screen "D_GraphicView_1" 800x480
   GraphicView "Static" at 6,4 size 100x60
   TextField "Label_Static" at 6,96 size 148x16; Text 'Static'
   GraphicView "A_Range" at 158,4 size 100x60
      Appearance <- "D_Range"
   TextField "Label_A_Range" at 158,96 size 148x16; Text 'A_Range'
   GraphicView "A_Flash" at 310,4 size 100x60
      Appearance <- "D_Range"
   TextField "Label_A_Flash" at 310,96 size 148x16; Text 'A_Flash'
   GraphicView "A_Bit" at 462,4 size 100x60
      Appearance <- "D_Bool"
   TextField "Label_A_Bit" at 462,96 size 148x16; Text 'A_Bit'
   GraphicView "A_Bits" at 614,4 size 100x60
      Appearance <- "D_Bits"
   TextField "Label_A_Bits" at 614,96 size 148x16; Text 'A_Bits'
   GraphicView "V_Range" at 6,116 size 100x60
      Visibility <- "D_Range"
   TextField "Label_V_Range" at 6,208 size 148x16; Text 'V_Range'
   GraphicView "V_Bit" at 158,116 size 100x60
      Visibility <- "D_Vis"
   TextField "Label_V_Bit" at 158,208 size 148x16; Text 'V_Bit'
   GraphicView "M_H" at 310,116 size 100x60
      HorizontalMovement <- "D_Pct"
   TextField "Label_M_H" at 310,208 size 148x16; Text 'M_H'
   GraphicView "M_V" at 462,116 size 100x60
      VerticalMovement <- "D_Pct"
   TextField "Label_M_V" at 462,208 size 148x16; Text 'M_V'
   GraphicView "M_D" at 614,116 size 100x60
      DiagonalMovement <- "D_Pct"
   TextField "Label_M_D" at 614,208 size 148x16; Text 'M_D'
   GraphicView "M_Direct" at 6,228 size 100x60
      DirectMovement <- "D_X"
      DirectMovement <- "D_Y"
   TextField "Label_M_Direct" at 6,320 size 148x16; Text 'M_Direct'
   GraphicView "E_Range" at 158,228 size 100x60
      ObjectEnable <- "D_Range"
   TextField "Label_E_Range" at 158,320 size 148x16; Text 'E_Range'
   GraphicView "E_Bit" at 310,228 size 100x60
      ObjectEnable <- "D_En"
   TextField "Label_E_Bit" at 310,320 size 148x16; Text 'E_Bit'
   IOField "State" at 4,454 size 60x22; FormatPattern 9
      ProcessValue <- "D_State"
   Button "S1" at 70,454 size 40x22; TextOff 'S1'
      on Click: "SetS1"()
   Button "S2" at 114,454 size 40x22; TextOff 'S2'
      on Click: "SetS2"()
   Button "S3" at 158,454 size 40x22; TextOff 'S3'
      on Click: "SetS3"()
   Button "S4" at 202,454 size 40x22; TextOff 'S4'
      on Click: "SetS4"()
   Button "Next" at 756,454 size 40x22; TextOff 'Next'
      on Click: ActivateScreen("D_IOField_1", 0)

screen "D_IOField_2" 800x480
   IOField "PV_Int_Output" at 6,4 size 100x30; FormatPattern s99999
      ProcessValue <- "D_Int"
   TextField "Label_PV_Int_Output" at 6,66 size 148x16; Text 'PV_Int_Output'
   IOField "PV_Int_s99" at 158,4 size 100x30; FormatPattern s99
      ProcessValue <- "D_Int"
   TextField "Label_PV_Int_s99" at 158,66 size 148x16; Text 'PV_Int_s99'
   IOField "State" at 4,454 size 60x22; FormatPattern 9
      ProcessValue <- "D_State"
   Button "S1" at 70,454 size 40x22; TextOff 'S1'
      on Click: "SetS1"()
   Button "S2" at 114,454 size 40x22; TextOff 'S2'
      on Click: "SetS2"()
   Button "S3" at 158,454 size 40x22; TextOff 'S3'
      on Click: "SetS3"()
   Button "S4" at 202,454 size 40x22; TextOff 'S4'
      on Click: "SetS4"()
   Button "Next" at 756,454 size 40x22; TextOff 'Next'
      on Click: ActivateScreen("D_Button_1", 0)

screen "D_Line_1" 800x480
   TextField "Label_Static" at 6,86 size 148x16; Text 'Static'
   Line "A_Range" at 158,4 size 100x50
      Appearance <- "D_Range"
   TextField "Label_A_Range" at 158,86 size 148x16; Text 'A_Range'
   Line "A_Flash" at 310,4 size 100x50
      Appearance <- "D_Range"
   TextField "Label_A_Flash" at 310,86 size 148x16; Text 'A_Flash'
   Line "A_Bit" at 462,4 size 100x50
      Appearance <- "D_Bool"
   TextField "Label_A_Bit" at 462,86 size 148x16; Text 'A_Bit'
   Line "A_Bits" at 614,4 size 100x50
      Appearance <- "D_Bits"
   TextField "Label_A_Bits" at 614,86 size 148x16; Text 'A_Bits'
   Line "V_Range" at 6,106 size 100x50
      Visibility <- "D_Range"
   TextField "Label_V_Range" at 6,188 size 148x16; Text 'V_Range'
   Line "V_Bit" at 158,106 size 100x50
      Visibility <- "D_Vis"
   TextField "Label_V_Bit" at 158,188 size 148x16; Text 'V_Bit'
   Line "M_H" at 310,106 size 100x50
      HorizontalMovement <- "D_Pct"
   TextField "Label_M_H" at 310,188 size 148x16; Text 'M_H'
   Line "M_V" at 462,106 size 100x50
      VerticalMovement <- "D_Pct"
   TextField "Label_M_V" at 462,188 size 148x16; Text 'M_V'
   Line "M_D" at 614,106 size 100x50
      DiagonalMovement <- "D_Pct"
   TextField "Label_M_D" at 614,188 size 148x16; Text 'M_D'
   Line "M_Direct" at 6,208 size 100x50
      DirectMovement <- "D_X"
      DirectMovement <- "D_Y"
   TextField "Label_M_Direct" at 6,290 size 148x16; Text 'M_Direct'
   Line "E_Range" at 158,208 size 100x50
      ObjectEnable <- "D_Range"
   TextField "Label_E_Range" at 158,290 size 148x16; Text 'E_Range'
   Line "E_Bit" at 310,208 size 100x50
      ObjectEnable <- "D_En"
   TextField "Label_E_Bit" at 310,290 size 148x16; Text 'E_Bit'
   IOField "State" at 4,454 size 60x22; FormatPattern 9
      ProcessValue <- "D_State"
   Button "S1" at 70,454 size 40x22; TextOff 'S1'
      on Click: "SetS1"()
   Button "S2" at 114,454 size 40x22; TextOff 'S2'
      on Click: "SetS2"()
   Button "S3" at 158,454 size 40x22; TextOff 'S3'
      on Click: "SetS3"()
   Button "S4" at 202,454 size 40x22; TextOff 'S4'
      on Click: "SetS4"()
   Button "Next" at 756,454 size 40x22; TextOff 'Next'
      on Click: ActivateScreen("D_Polyline_1", 0)

screen "D_Polygon_1" 800x480
   TextField "Label_Static" at 6,86 size 148x16; Text 'Static'
   Polygon "A_Range" at 158,4 size 100x50
      Appearance <- "D_Range"
   TextField "Label_A_Range" at 158,86 size 148x16; Text 'A_Range'
   Polygon "A_Flash" at 310,4 size 100x50
      Appearance <- "D_Range"
   TextField "Label_A_Flash" at 310,86 size 148x16; Text 'A_Flash'
   Polygon "A_Bit" at 462,4 size 100x50
      Appearance <- "D_Bool"
   TextField "Label_A_Bit" at 462,86 size 148x16; Text 'A_Bit'
   Polygon "A_Bits" at 614,4 size 100x50
      Appearance <- "D_Bits"
   TextField "Label_A_Bits" at 614,86 size 148x16; Text 'A_Bits'
   Polygon "V_Range" at 6,106 size 100x50
      Visibility <- "D_Range"
   TextField "Label_V_Range" at 6,188 size 148x16; Text 'V_Range'
   Polygon "V_Bit" at 158,106 size 100x50
      Visibility <- "D_Vis"
   TextField "Label_V_Bit" at 158,188 size 148x16; Text 'V_Bit'
   Polygon "M_H" at 310,106 size 100x50
      HorizontalMovement <- "D_Pct"
   TextField "Label_M_H" at 310,188 size 148x16; Text 'M_H'
   Polygon "M_V" at 462,106 size 100x50
      VerticalMovement <- "D_Pct"
   TextField "Label_M_V" at 462,188 size 148x16; Text 'M_V'
   Polygon "M_D" at 614,106 size 100x50
      DiagonalMovement <- "D_Pct"
   TextField "Label_M_D" at 614,188 size 148x16; Text 'M_D'
   Polygon "M_Direct" at 6,208 size 100x50
      DirectMovement <- "D_X"
      DirectMovement <- "D_Y"
   TextField "Label_M_Direct" at 6,290 size 148x16; Text 'M_Direct'
   Polygon "E_Range" at 158,208 size 100x50
      ObjectEnable <- "D_Range"
   TextField "Label_E_Range" at 158,290 size 148x16; Text 'E_Range'
   Polygon "E_Bit" at 310,208 size 100x50
      ObjectEnable <- "D_En"
   TextField "Label_E_Bit" at 310,290 size 148x16; Text 'E_Bit'
   IOField "State" at 4,454 size 60x22; FormatPattern 9
      ProcessValue <- "D_State"
   Button "S1" at 70,454 size 40x22; TextOff 'S1'
      on Click: "SetS1"()
   Button "S2" at 114,454 size 40x22; TextOff 'S2'
      on Click: "SetS2"()
   Button "S3" at 158,454 size 40x22; TextOff 'S3'
      on Click: "SetS3"()
   Button "S4" at 202,454 size 40x22; TextOff 'S4'
      on Click: "SetS4"()
   Button "Next" at 756,454 size 40x22; TextOff 'Next'
      on Click: ActivateScreen("D_Ellipse_1", 0)

screen "D_Polyline_1" 800x480
   TextField "Label_Static" at 6,86 size 148x16; Text 'Static'
   Polyline "A_Range" at 158,4 size 100x50
      Appearance <- "D_Range"
   TextField "Label_A_Range" at 158,86 size 148x16; Text 'A_Range'
   Polyline "A_Flash" at 310,4 size 100x50
      Appearance <- "D_Range"
   TextField "Label_A_Flash" at 310,86 size 148x16; Text 'A_Flash'
   Polyline "A_Bit" at 462,4 size 100x50
      Appearance <- "D_Bool"
   TextField "Label_A_Bit" at 462,86 size 148x16; Text 'A_Bit'
   Polyline "A_Bits" at 614,4 size 100x50
      Appearance <- "D_Bits"
   TextField "Label_A_Bits" at 614,86 size 148x16; Text 'A_Bits'
   Polyline "V_Range" at 6,106 size 100x50
      Visibility <- "D_Range"
   TextField "Label_V_Range" at 6,188 size 148x16; Text 'V_Range'
   Polyline "V_Bit" at 158,106 size 100x50
      Visibility <- "D_Vis"
   TextField "Label_V_Bit" at 158,188 size 148x16; Text 'V_Bit'
   Polyline "M_H" at 310,106 size 100x50
      HorizontalMovement <- "D_Pct"
   TextField "Label_M_H" at 310,188 size 148x16; Text 'M_H'
   Polyline "M_V" at 462,106 size 100x50
      VerticalMovement <- "D_Pct"
   TextField "Label_M_V" at 462,188 size 148x16; Text 'M_V'
   Polyline "M_D" at 614,106 size 100x50
      DiagonalMovement <- "D_Pct"
   TextField "Label_M_D" at 614,188 size 148x16; Text 'M_D'
   Polyline "M_Direct" at 6,208 size 100x50
      DirectMovement <- "D_X"
      DirectMovement <- "D_Y"
   TextField "Label_M_Direct" at 6,290 size 148x16; Text 'M_Direct'
   Polyline "E_Range" at 158,208 size 100x50
      ObjectEnable <- "D_Range"
   TextField "Label_E_Range" at 158,290 size 148x16; Text 'E_Range'
   Polyline "E_Bit" at 310,208 size 100x50
      ObjectEnable <- "D_En"
   TextField "Label_E_Bit" at 310,290 size 148x16; Text 'E_Bit'
   IOField "State" at 4,454 size 60x22; FormatPattern 9
      ProcessValue <- "D_State"
   Button "S1" at 70,454 size 40x22; TextOff 'S1'
      on Click: "SetS1"()
   Button "S2" at 114,454 size 40x22; TextOff 'S2'
      on Click: "SetS2"()
   Button "S3" at 158,454 size 40x22; TextOff 'S3'
      on Click: "SetS3"()
   Button "S4" at 202,454 size 40x22; TextOff 'S4'
      on Click: "SetS4"()
   Button "Next" at 756,454 size 40x22; TextOff 'Next'
      on Click: ActivateScreen("D_Polygon_1", 0)

screen "D_Rectangle_1" 800x480
   TextField "Label_Static" at 6,86 size 148x16; Text 'Static'
   Rectangle "A_Range" at 158,4 size 100x50
      Appearance <- "D_Range"
   TextField "Label_A_Range" at 158,86 size 148x16; Text 'A_Range'
   Rectangle "A_Flash" at 310,4 size 100x50
      Appearance <- "D_Range"
   TextField "Label_A_Flash" at 310,86 size 148x16; Text 'A_Flash'
   Rectangle "A_Bit" at 462,4 size 100x50
      Appearance <- "D_Bool"
   TextField "Label_A_Bit" at 462,86 size 148x16; Text 'A_Bit'
   Rectangle "A_Bits" at 614,4 size 100x50
      Appearance <- "D_Bits"
   TextField "Label_A_Bits" at 614,86 size 148x16; Text 'A_Bits'
   Rectangle "V_Range" at 6,106 size 100x50
      Visibility <- "D_Range"
   TextField "Label_V_Range" at 6,188 size 148x16; Text 'V_Range'
   Rectangle "V_Bit" at 158,106 size 100x50
      Visibility <- "D_Vis"
   TextField "Label_V_Bit" at 158,188 size 148x16; Text 'V_Bit'
   Rectangle "M_H" at 310,106 size 100x50
      HorizontalMovement <- "D_Pct"
   TextField "Label_M_H" at 310,188 size 148x16; Text 'M_H'
   Rectangle "M_V" at 462,106 size 100x50
      VerticalMovement <- "D_Pct"
   TextField "Label_M_V" at 462,188 size 148x16; Text 'M_V'
   Rectangle "M_D" at 614,106 size 100x50
      DiagonalMovement <- "D_Pct"
   TextField "Label_M_D" at 614,188 size 148x16; Text 'M_D'
   Rectangle "M_Direct" at 6,208 size 100x50
      DirectMovement <- "D_X"
      DirectMovement <- "D_Y"
   TextField "Label_M_Direct" at 6,290 size 148x16; Text 'M_Direct'
   Rectangle "E_Range" at 158,208 size 100x50
      ObjectEnable <- "D_Range"
   TextField "Label_E_Range" at 158,290 size 148x16; Text 'E_Range'
   Rectangle "E_Bit" at 310,208 size 100x50
      ObjectEnable <- "D_En"
   TextField "Label_E_Bit" at 310,290 size 148x16; Text 'E_Bit'
   IOField "State" at 4,454 size 60x22; FormatPattern 9
      ProcessValue <- "D_State"
   Button "S1" at 70,454 size 40x22; TextOff 'S1'
      on Click: "SetS1"()
   Button "S2" at 114,454 size 40x22; TextOff 'S2'
      on Click: "SetS2"()
   Button "S3" at 158,454 size 40x22; TextOff 'S3'
      on Click: "SetS3"()
   Button "S4" at 202,454 size 40x22; TextOff 'S4'
      on Click: "SetS4"()
   Button "Next" at 756,454 size 40x22; TextOff 'Next'
      on Click: ActivateScreen("D_TextField_1", 0)

screen "D_Switch_1" 800x480
   Switch "Static" at 6,4 size 120x40; CaptionText 'Switch'; TextOff '0'; TextOn '1'
   TextField "Label_Static" at 6,76 size 168x16; Text 'Static'
   Switch "A_Range" at 178,4 size 120x40; CaptionText 'Switch'; TextOff '0'; TextOn '1'
      Appearance <- "D_Range"
   TextField "Label_A_Range" at 178,76 size 168x16; Text 'A_Range'
   Switch "A_Flash" at 350,4 size 120x40; CaptionText 'Switch'; TextOff '0'; TextOn '1'
      Appearance <- "D_Range"
   TextField "Label_A_Flash" at 350,76 size 168x16; Text 'A_Flash'
   Switch "A_Bit" at 522,4 size 120x40; CaptionText 'Switch'; TextOff '0'; TextOn '1'
      Appearance <- "D_Bool"
   TextField "Label_A_Bit" at 522,76 size 168x16; Text 'A_Bit'
   Switch "A_Bits" at 6,96 size 120x40; CaptionText 'Switch'; TextOff '0'; TextOn '1'
      Appearance <- "D_Bits"
   TextField "Label_A_Bits" at 6,168 size 168x16; Text 'A_Bits'
   Switch "V_Range" at 178,96 size 120x40; CaptionText 'Switch'; TextOff '0'; TextOn '1'
      Visibility <- "D_Range"
   TextField "Label_V_Range" at 178,168 size 168x16; Text 'V_Range'
   Switch "V_Bit" at 350,96 size 120x40; CaptionText 'Switch'; TextOff '0'; TextOn '1'
      Visibility <- "D_Vis"
   TextField "Label_V_Bit" at 350,168 size 168x16; Text 'V_Bit'
   Switch "M_H" at 522,96 size 120x40; CaptionText 'Switch'; TextOff '0'; TextOn '1'
      HorizontalMovement <- "D_Pct"
   TextField "Label_M_H" at 522,168 size 168x16; Text 'M_H'
   Switch "M_V" at 6,188 size 120x40; CaptionText 'Switch'; TextOff '0'; TextOn '1'
      VerticalMovement <- "D_Pct"
   TextField "Label_M_V" at 6,260 size 168x16; Text 'M_V'
   Switch "M_D" at 178,188 size 120x40; CaptionText 'Switch'; TextOff '0'; TextOn '1'
      DiagonalMovement <- "D_Pct"
   TextField "Label_M_D" at 178,260 size 168x16; Text 'M_D'
   Switch "M_Direct" at 350,188 size 120x40; CaptionText 'Switch'; TextOff '0'; TextOn '1'
      DirectMovement <- "D_X"
      DirectMovement <- "D_Y"
   TextField "Label_M_Direct" at 350,260 size 168x16; Text 'M_Direct'
   Switch "E_Range" at 522,188 size 120x40; CaptionText 'Switch'; TextOff '0'; TextOn '1'
      ObjectEnable <- "D_Range"
   TextField "Label_E_Range" at 522,260 size 168x16; Text 'E_Range'
   Switch "E_Bit" at 6,280 size 120x40; CaptionText 'Switch'; TextOff '0'; TextOn '1'
      ObjectEnable <- "D_En"
   TextField "Label_E_Bit" at 6,352 size 168x16; Text 'E_Bit'
   Switch "PV_Bool" at 178,280 size 120x40; CaptionText 'Switch'; TextOff '0'; TextOn '1'
      ProcessValue <- "D_Bool"
   TextField "Label_PV_Bool" at 178,352 size 168x16; Text 'PV_Bool'
   IOField "State" at 4,454 size 60x22; FormatPattern 9
      ProcessValue <- "D_State"
   Button "S1" at 70,454 size 40x22; TextOff 'S1'
      on Click: "SetS1"()
   Button "S2" at 114,454 size 40x22; TextOff 'S2'
      on Click: "SetS2"()
   Button "S3" at 158,454 size 40x22; TextOff 'S3'
      on Click: "SetS3"()
   Button "S4" at 202,454 size 40x22; TextOff 'S4'
      on Click: "SetS4"()
   Button "Next" at 756,454 size 40x22; TextOff 'Next'
      on Click: ActivateScreen("D_SymbolLibrary_1", 0)

screen "D_SymbolicIOField_1" 800x480
   SymbolicIOField "Static" at 6,4 size 120x30; TextOff '0'; TextOn '1'
   TextField "Label_Static" at 6,66 size 168x16; Text 'Static'
   SymbolicIOField "A_Range" at 178,4 size 120x30; TextOff '0'; TextOn '1'
      Appearance <- "D_Range"
   TextField "Label_A_Range" at 178,66 size 168x16; Text 'A_Range'
   SymbolicIOField "A_Flash" at 350,4 size 120x30; TextOff '0'; TextOn '1'
      Appearance <- "D_Range"
   TextField "Label_A_Flash" at 350,66 size 168x16; Text 'A_Flash'
   SymbolicIOField "A_Bit" at 522,4 size 120x30; TextOff '0'; TextOn '1'
      Appearance <- "D_Bool"
   TextField "Label_A_Bit" at 522,66 size 168x16; Text 'A_Bit'
   SymbolicIOField "A_Bits" at 6,86 size 120x30; TextOff '0'; TextOn '1'
      Appearance <- "D_Bits"
   TextField "Label_A_Bits" at 6,148 size 168x16; Text 'A_Bits'
   SymbolicIOField "V_Range" at 178,86 size 120x30; TextOff '0'; TextOn '1'
      Visibility <- "D_Range"
   TextField "Label_V_Range" at 178,148 size 168x16; Text 'V_Range'
   SymbolicIOField "V_Bit" at 350,86 size 120x30; TextOff '0'; TextOn '1'
      Visibility <- "D_Vis"
   TextField "Label_V_Bit" at 350,148 size 168x16; Text 'V_Bit'
   SymbolicIOField "M_H" at 522,86 size 120x30; TextOff '0'; TextOn '1'
      HorizontalMovement <- "D_Pct"
   TextField "Label_M_H" at 522,148 size 168x16; Text 'M_H'
   SymbolicIOField "M_V" at 6,168 size 120x30; TextOff '0'; TextOn '1'
      VerticalMovement <- "D_Pct"
   TextField "Label_M_V" at 6,230 size 168x16; Text 'M_V'
   SymbolicIOField "M_D" at 178,168 size 120x30; TextOff '0'; TextOn '1'
      DiagonalMovement <- "D_Pct"
   TextField "Label_M_D" at 178,230 size 168x16; Text 'M_D'
   SymbolicIOField "M_Direct" at 350,168 size 120x30; TextOff '0'; TextOn '1'
      DirectMovement <- "D_X"
      DirectMovement <- "D_Y"
   TextField "Label_M_Direct" at 350,230 size 168x16; Text 'M_Direct'
   SymbolicIOField "E_Range" at 522,168 size 120x30; TextOff '0'; TextOn '1'
      ObjectEnable <- "D_Range"
   TextField "Label_E_Range" at 522,230 size 168x16; Text 'E_Range'
   SymbolicIOField "E_Bit" at 6,250 size 120x30; TextOff '0'; TextOn '1'
      ObjectEnable <- "D_En"
   TextField "Label_E_Bit" at 6,312 size 168x16; Text 'E_Bit'
   SymbolicIOField "PV_TL_Value" at 178,250 size 120x30; TextOff '0'; TextOn '1'; TextList "TL_Value"
      ProcessValue <- "D_TL"
   TextField "Label_PV_TL_Value" at 178,312 size 168x16; Text 'PV_TL_Value'
   SymbolicIOField "PV_TL_Bit" at 350,250 size 120x30; TextOff '0'; TextOn '1'; TextList "TL_Bit"
      ProcessValue <- "D_Bool"
   TextField "Label_PV_TL_Bit" at 350,312 size 168x16; Text 'PV_TL_Bit'
   SymbolicIOField "PV_TL_BitNo" at 522,250 size 120x30; TextOff '0'; TextOn '1'; TextList "TL_BitNo"
      ProcessValue <- "D_Bits"
   TextField "Label_PV_TL_BitNo" at 522,312 size 168x16; Text 'PV_TL_BitNo'
   IOField "State" at 4,454 size 60x22; FormatPattern 9
      ProcessValue <- "D_State"
   Button "S1" at 70,454 size 40x22; TextOff 'S1'
      on Click: "SetS1"()
   Button "S2" at 114,454 size 40x22; TextOff 'S2'
      on Click: "SetS2"()
   Button "S3" at 158,454 size 40x22; TextOff 'S3'
      on Click: "SetS3"()
   Button "S4" at 202,454 size 40x22; TextOff 'S4'
      on Click: "SetS4"()
   Button "Next" at 756,454 size 40x22; TextOff 'Next'
      on Click: ActivateScreen("D_GraphicIOField_1", 0)

screen "D_TextField_1" 800x480
   TextField "Static" at 6,4 size 100x30; Text 'Text'
   TextField "Label_Static" at 6,66 size 148x16; Text 'Static'
   TextField "A_Range" at 158,4 size 100x30; Text 'Text'
      Appearance <- "D_Range"
   TextField "Label_A_Range" at 158,66 size 148x16; Text 'A_Range'
   TextField "A_Flash" at 310,4 size 100x30; Text 'Text'
      Appearance <- "D_Range"
   TextField "Label_A_Flash" at 310,66 size 148x16; Text 'A_Flash'
   TextField "A_Bit" at 462,4 size 100x30; Text 'Text'
      Appearance <- "D_Bool"
   TextField "Label_A_Bit" at 462,66 size 148x16; Text 'A_Bit'
   TextField "A_Bits" at 614,4 size 100x30; Text 'Text'
      Appearance <- "D_Bits"
   TextField "Label_A_Bits" at 614,66 size 148x16; Text 'A_Bits'
   TextField "V_Range" at 6,86 size 100x30; Text 'Text'
      Visibility <- "D_Range"
   TextField "Label_V_Range" at 6,148 size 148x16; Text 'V_Range'
   TextField "V_Bit" at 158,86 size 100x30; Text 'Text'
      Visibility <- "D_Vis"
   TextField "Label_V_Bit" at 158,148 size 148x16; Text 'V_Bit'
   TextField "M_H" at 310,86 size 100x30; Text 'Text'
      HorizontalMovement <- "D_Pct"
   TextField "Label_M_H" at 310,148 size 148x16; Text 'M_H'
   TextField "M_V" at 462,86 size 100x30; Text 'Text'
      VerticalMovement <- "D_Pct"
   TextField "Label_M_V" at 462,148 size 148x16; Text 'M_V'
   TextField "M_D" at 614,86 size 100x30; Text 'Text'
      DiagonalMovement <- "D_Pct"
   TextField "Label_M_D" at 614,148 size 148x16; Text 'M_D'
   TextField "M_Direct" at 6,168 size 100x30; Text 'Text'
      DirectMovement <- "D_X"
      DirectMovement <- "D_Y"
   TextField "Label_M_Direct" at 6,230 size 148x16; Text 'M_Direct'
   TextField "E_Range" at 158,168 size 100x30; Text 'Text'
      ObjectEnable <- "D_Range"
   TextField "Label_E_Range" at 158,230 size 148x16; Text 'E_Range'
   TextField "E_Bit" at 310,168 size 100x30; Text 'Text'
      ObjectEnable <- "D_En"
   TextField "Label_E_Bit" at 310,230 size 148x16; Text 'E_Bit'
   IOField "State" at 4,454 size 60x22; FormatPattern 9
      ProcessValue <- "D_State"
   Button "S1" at 70,454 size 40x22; TextOff 'S1'
      on Click: "SetS1"()
   Button "S2" at 114,454 size 40x22; TextOff 'S2'
      on Click: "SetS2"()
   Button "S3" at 158,454 size 40x22; TextOff 'S3'
      on Click: "SetS3"()
   Button "S4" at 202,454 size 40x22; TextOff 'S4'
      on Click: "SetS4"()
   Button "Next" at 756,454 size 40x22; TextOff 'Next'
      on Click: ActivateScreen("D_GraphicView_1", 0)

screen "D_IOField_1" 800x480
   IOField "Static" at 6,4 size 100x30
   TextField "Label_Static" at 6,66 size 148x16; Text 'Static'
   IOField "A_Range" at 158,4 size 100x30
      Appearance <- "D_Range"
   TextField "Label_A_Range" at 158,66 size 148x16; Text 'A_Range'
   IOField "A_Flash" at 310,4 size 100x30
      Appearance <- "D_Range"
   TextField "Label_A_Flash" at 310,66 size 148x16; Text 'A_Flash'
   IOField "A_Bit" at 462,4 size 100x30
      Appearance <- "D_Bool"
   TextField "Label_A_Bit" at 462,66 size 148x16; Text 'A_Bit'
   IOField "A_Bits" at 614,4 size 100x30
      Appearance <- "D_Bits"
   TextField "Label_A_Bits" at 614,66 size 148x16; Text 'A_Bits'
   IOField "V_Range" at 6,86 size 100x30
      Visibility <- "D_Range"
   TextField "Label_V_Range" at 6,148 size 148x16; Text 'V_Range'
   IOField "V_Bit" at 158,86 size 100x30
      Visibility <- "D_Vis"
   TextField "Label_V_Bit" at 158,148 size 148x16; Text 'V_Bit'
   IOField "M_H" at 310,86 size 100x30
      HorizontalMovement <- "D_Pct"
   TextField "Label_M_H" at 310,148 size 148x16; Text 'M_H'
   IOField "M_V" at 462,86 size 100x30
      VerticalMovement <- "D_Pct"
   TextField "Label_M_V" at 462,148 size 148x16; Text 'M_V'
   IOField "M_D" at 614,86 size 100x30
      DiagonalMovement <- "D_Pct"
   TextField "Label_M_D" at 614,148 size 148x16; Text 'M_D'
   IOField "M_Direct" at 6,168 size 100x30
      DirectMovement <- "D_X"
      DirectMovement <- "D_Y"
   TextField "Label_M_Direct" at 6,230 size 148x16; Text 'M_Direct'
   IOField "E_Range" at 158,168 size 100x30
      ObjectEnable <- "D_Range"
   TextField "Label_E_Range" at 158,230 size 148x16; Text 'E_Range'
   IOField "E_Bit" at 310,168 size 100x30
      ObjectEnable <- "D_En"
   TextField "Label_E_Bit" at 310,230 size 148x16; Text 'E_Bit'
   IOField "PV_SInt" at 462,168 size 100x30; FormatPattern s999
      ProcessValue <- "D_SInt"
   TextField "Label_PV_SInt" at 462,230 size 148x16; Text 'PV_SInt'
   IOField "PV_Int" at 614,168 size 100x30; FormatPattern s99999
      ProcessValue <- "D_Int"
   TextField "Label_PV_Int" at 614,230 size 148x16; Text 'PV_Int'
   IOField "PV_DInt" at 6,250 size 100x30; FormatPattern s9999999999
      ProcessValue <- "D_DInt"
   TextField "Label_PV_DInt" at 6,312 size 148x16; Text 'PV_DInt'
   IOField "PV_USInt" at 158,250 size 100x30; FormatPattern 999
      ProcessValue <- "D_USInt"
   TextField "Label_PV_USInt" at 158,312 size 148x16; Text 'PV_USInt'
   IOField "PV_UInt" at 310,250 size 100x30; FormatPattern 99999
      ProcessValue <- "D_UInt"
   TextField "Label_PV_UInt" at 310,312 size 148x16; Text 'PV_UInt'
   IOField "PV_UDInt" at 462,250 size 100x30; FormatPattern 9999999999
      ProcessValue <- "D_UDInt"
   TextField "Label_PV_UDInt" at 462,312 size 148x16; Text 'PV_UDInt'
   IOField "PV_Real" at 614,250 size 100x30
      ProcessValue <- "D_Real"
   TextField "Label_PV_Real" at 614,312 size 148x16; Text 'PV_Real'
   IOField "PV_LReal" at 6,332 size 100x30
      ProcessValue <- "D_LReal"
   TextField "Label_PV_LReal" at 6,394 size 148x16; Text 'PV_LReal'
   IOField "PV_String" at 158,332 size 100x30
      ProcessValue <- "D_String"
   TextField "Label_PV_String" at 158,394 size 148x16; Text 'PV_String'
   IOField "PV_Int_Shift2" at 310,332 size 100x30; FormatPattern s99999
      ProcessValue <- "D_Int"
   TextField "Label_PV_Int_Shift2" at 310,394 size 148x16; Text 'PV_Int_Shift2'
   IOField "PV_Int_s999999" at 462,332 size 100x30; FormatPattern s999999
      ProcessValue <- "D_Int"
   TextField "Label_PV_Int_s999999" at 462,394 size 148x16; Text 'PV_Int_s999999'
   IOField "PV_Real_s9999_99" at 614,332 size 100x30; FormatPattern s9999.99
      ProcessValue <- "D_Real"
   TextField "Label_PV_Real_s9999_99" at 614,394 size 148x16; Text 'PV_Real_s9999_99'
   IOField "State" at 4,454 size 60x22; FormatPattern 9
      ProcessValue <- "D_State"
   Button "S1" at 70,454 size 40x22; TextOff 'S1'
      on Click: "SetS1"()
   Button "S2" at 114,454 size 40x22; TextOff 'S2'
      on Click: "SetS2"()
   Button "S3" at 158,454 size 40x22; TextOff 'S3'
      on Click: "SetS3"()
   Button "S4" at 202,454 size 40x22; TextOff 'S4'
      on Click: "SetS4"()
   Button "Next" at 756,454 size 40x22; TextOff 'Next'
      on Click: ActivateScreen("D_IOField_2", 0)

screen "D_Bar_1" 800x480
   Bar "Static" at 6,4 size 40x120
   TextField "Label_Static" at 6,156 size 88x16; Text 'Static'
   Bar "A_Range" at 98,4 size 40x120
      Appearance <- "D_Range"
   TextField "Label_A_Range" at 98,156 size 88x16; Text 'A_Range'
   Bar "A_Flash" at 190,4 size 40x120
      Appearance <- "D_Range"
   TextField "Label_A_Flash" at 190,156 size 88x16; Text 'A_Flash'
   Bar "A_Bit" at 282,4 size 40x120
      Appearance <- "D_Bool"
   TextField "Label_A_Bit" at 282,156 size 88x16; Text 'A_Bit'
   Bar "A_Bits" at 374,4 size 40x120
      Appearance <- "D_Bits"
   TextField "Label_A_Bits" at 374,156 size 88x16; Text 'A_Bits'
   Bar "V_Range" at 466,4 size 40x120
      Visibility <- "D_Range"
   TextField "Label_V_Range" at 466,156 size 88x16; Text 'V_Range'
   Bar "V_Bit" at 558,4 size 40x120
      Visibility <- "D_Vis"
   TextField "Label_V_Bit" at 558,156 size 88x16; Text 'V_Bit'
   Bar "M_H" at 650,4 size 40x120
      HorizontalMovement <- "D_Pct"
   TextField "Label_M_H" at 650,156 size 88x16; Text 'M_H'
   Bar "M_V" at 6,176 size 40x120
      VerticalMovement <- "D_Pct"
   TextField "Label_M_V" at 6,328 size 88x16; Text 'M_V'
   Bar "M_D" at 98,176 size 40x120
      DiagonalMovement <- "D_Pct"
   TextField "Label_M_D" at 98,328 size 88x16; Text 'M_D'
   Bar "M_Direct" at 190,176 size 40x120
      DirectMovement <- "D_X"
      DirectMovement <- "D_Y"
   TextField "Label_M_Direct" at 190,328 size 88x16; Text 'M_Direct'
   Bar "E_Range" at 282,176 size 40x120
      ObjectEnable <- "D_Range"
   TextField "Label_E_Range" at 282,328 size 88x16; Text 'E_Range'
   Bar "E_Bit" at 374,176 size 40x120
      ObjectEnable <- "D_En"
   TextField "Label_E_Bit" at 374,328 size 88x16; Text 'E_Bit'
   Bar "PV_Pct" at 466,176 size 40x120
      ProcessValue <- "D_Pct"
   TextField "Label_PV_Pct" at 466,328 size 88x16; Text 'PV_Pct'
   Bar "PV_Real" at 558,176 size 40x120
      ProcessValue <- "D_Real"
   TextField "Label_PV_Real" at 558,328 size 88x16; Text 'PV_Real'
   Bar "PV_BarR" at 650,176 size 40x120
      ProcessValue <- "D_BarR"
   TextField "Label_PV_BarR" at 650,328 size 88x16; Text 'PV_BarR'
   IOField "State" at 4,454 size 60x22; FormatPattern 9
      ProcessValue <- "D_State"
   Button "S1" at 70,454 size 40x22; TextOff 'S1'
      on Click: "SetS1"()
   Button "S2" at 114,454 size 40x22; TextOff 'S2'
      on Click: "SetS2"()
   Button "S3" at 158,454 size 40x22; TextOff 'S3'
      on Click: "SetS3"()
   Button "S4" at 202,454 size 40x22; TextOff 'S4'
      on Click: "SetS4"()
   Button "Next" at 756,454 size 40x22; TextOff 'Next'
      on Click: ActivateScreen("D_Bar_2", 0)

screen "D_Bar_2" 800x480
   Bar "PV_Pct_0_100" at 6,4 size 40x120; MinimumValue 0; MaximumValue 100
      ProcessValue <- "D_Pct"
   TextField "Label_PV_Pct_0_100" at 6,156 size 88x16; Text 'PV_Pct_0_100'
   Bar "PV_Pct_MaxMin" at 98,4 size 40x120
      ProcessValue <- "D_Pct"
      MaximumValue <- "D_Max"
      MinimumValue <- "D_Min"
   TextField "Label_PV_Pct_MaxMin" at 98,156 size 88x16; Text 'PV_Pct_MaxMin'
   IOField "State" at 4,454 size 60x22; FormatPattern 9
      ProcessValue <- "D_State"
   Button "S1" at 70,454 size 40x22; TextOff 'S1'
      on Click: "SetS1"()
   Button "S2" at 114,454 size 40x22; TextOff 'S2'
      on Click: "SetS2"()
   Button "S3" at 158,454 size 40x22; TextOff 'S3'
      on Click: "SetS3"()
   Button "S4" at 202,454 size 40x22; TextOff 'S4'
      on Click: "SetS4"()
   Button "Next" at 756,454 size 40x22; TextOff 'Next'
      on Click: ActivateScreen("D_Switch_1", 0)

screen "D_Gauge_1" 800x480
   Gauge "Static" at 6,4 size 150x150; CaptionText 'SIMATIC'
   TextField "Label_Static" at 6,186 size 198x16; Text 'Static'
   Gauge "A_Range" at 208,4 size 150x150; CaptionText 'SIMATIC'
      Appearance <- "D_Range"
   TextField "Label_A_Range" at 208,186 size 198x16; Text 'A_Range'
   Gauge "A_Flash" at 410,4 size 150x150; CaptionText 'SIMATIC'
      Appearance <- "D_Range"
   TextField "Label_A_Flash" at 410,186 size 198x16; Text 'A_Flash'
   Gauge "A_Bit" at 6,206 size 150x150; CaptionText 'SIMATIC'
      Appearance <- "D_Bool"
   TextField "Label_A_Bit" at 6,388 size 198x16; Text 'A_Bit'
   Gauge "A_Bits" at 208,206 size 150x150; CaptionText 'SIMATIC'
      Appearance <- "D_Bits"
   TextField "Label_A_Bits" at 208,388 size 198x16; Text 'A_Bits'
   Gauge "V_Range" at 410,206 size 150x150; CaptionText 'SIMATIC'
      Visibility <- "D_Range"
   TextField "Label_V_Range" at 410,388 size 198x16; Text 'V_Range'
   IOField "State" at 4,454 size 60x22; FormatPattern 9
      ProcessValue <- "D_State"
   Button "S1" at 70,454 size 40x22; TextOff 'S1'
      on Click: "SetS1"()
   Button "S2" at 114,454 size 40x22; TextOff 'S2'
      on Click: "SetS2"()
   Button "S3" at 158,454 size 40x22; TextOff 'S3'
      on Click: "SetS3"()
   Button "S4" at 202,454 size 40x22; TextOff 'S4'
      on Click: "SetS4"()
   Button "Next" at 756,454 size 40x22; TextOff 'Next'
      on Click: ActivateScreen("D_Gauge_2", 0)

screen "D_Gauge_2" 800x480
   Gauge "V_Bit" at 6,4 size 150x150; CaptionText 'SIMATIC'
      Visibility <- "D_Vis"
   TextField "Label_V_Bit" at 6,186 size 198x16; Text 'V_Bit'
   Gauge "M_H" at 208,4 size 150x150; CaptionText 'SIMATIC'
      HorizontalMovement <- "D_Pct"
   TextField "Label_M_H" at 208,186 size 198x16; Text 'M_H'
   Gauge "M_V" at 410,4 size 150x150; CaptionText 'SIMATIC'
      VerticalMovement <- "D_Pct"
   TextField "Label_M_V" at 410,186 size 198x16; Text 'M_V'
   Gauge "M_D" at 6,206 size 150x150; CaptionText 'SIMATIC'
      DiagonalMovement <- "D_Pct"
   TextField "Label_M_D" at 6,388 size 198x16; Text 'M_D'
   Gauge "M_Direct" at 208,206 size 150x150; CaptionText 'SIMATIC'
      DirectMovement <- "D_X"
      DirectMovement <- "D_Y"
   TextField "Label_M_Direct" at 208,388 size 198x16; Text 'M_Direct'
   Gauge "E_Range" at 410,206 size 150x150; CaptionText 'SIMATIC'
      ObjectEnable <- "D_Range"
   TextField "Label_E_Range" at 410,388 size 198x16; Text 'E_Range'
   IOField "State" at 4,454 size 60x22; FormatPattern 9
      ProcessValue <- "D_State"
   Button "S1" at 70,454 size 40x22; TextOff 'S1'
      on Click: "SetS1"()
   Button "S2" at 114,454 size 40x22; TextOff 'S2'
      on Click: "SetS2"()
   Button "S3" at 158,454 size 40x22; TextOff 'S3'
      on Click: "SetS3"()
   Button "S4" at 202,454 size 40x22; TextOff 'S4'
      on Click: "SetS4"()
   Button "Next" at 756,454 size 40x22; TextOff 'Next'
      on Click: ActivateScreen("D_Gauge_3", 0)

screen "D_Gauge_3" 800x480
   Gauge "E_Bit" at 6,4 size 150x150; CaptionText 'SIMATIC'
      ObjectEnable <- "D_En"
   TextField "Label_E_Bit" at 6,186 size 198x16; Text 'E_Bit'
   Gauge "PV_Pct" at 208,4 size 150x150; CaptionText 'SIMATIC'
      ProcessValue <- "D_Pct"
   TextField "Label_PV_Pct" at 208,186 size 198x16; Text 'PV_Pct'
   Gauge "PV_Real" at 410,4 size 150x150; CaptionText 'SIMATIC'
      ProcessValue <- "D_Real"
   TextField "Label_PV_Real" at 410,186 size 198x16; Text 'PV_Real'
   Gauge "PV_Pct_MaxMin" at 6,206 size 150x150; CaptionText 'SIMATIC'
      ProcessValue <- "D_Pct"
      MaximumValue <- "D_Max"
      MinimumValue <- "D_Min"
   TextField "Label_PV_Pct_MaxMin" at 6,388 size 198x16; Text 'PV_Pct_MaxMin'
   IOField "State" at 4,454 size 60x22; FormatPattern 9
      ProcessValue <- "D_State"
   Button "S1" at 70,454 size 40x22; TextOff 'S1'
      on Click: "SetS1"()
   Button "S2" at 114,454 size 40x22; TextOff 'S2'
      on Click: "SetS2"()
   Button "S3" at 158,454 size 40x22; TextOff 'S3'
      on Click: "SetS3"()
   Button "S4" at 202,454 size 40x22; TextOff 'S4'
      on Click: "SetS4"()
   Button "Next" at 756,454 size 40x22; TextOff 'Next'
      on Click: ActivateScreen("D_Clock_1", 0)

screen "D_Slider_1" 800x480
   Slider "Static" at 6,4 size 60x160; Caption 'SIMATIC'
   TextField "Label_Static" at 6,196 size 108x16; Text 'Static'
   Slider "A_Range" at 118,4 size 60x160; Caption 'SIMATIC'
      Appearance <- "D_Range"
   TextField "Label_A_Range" at 118,196 size 108x16; Text 'A_Range'
   Slider "A_Flash" at 230,4 size 60x160; Caption 'SIMATIC'
      Appearance <- "D_Range"
   TextField "Label_A_Flash" at 230,196 size 108x16; Text 'A_Flash'
   Slider "A_Bit" at 342,4 size 60x160; Caption 'SIMATIC'
      Appearance <- "D_Bool"
   TextField "Label_A_Bit" at 342,196 size 108x16; Text 'A_Bit'
   Slider "A_Bits" at 454,4 size 60x160; Caption 'SIMATIC'
      Appearance <- "D_Bits"
   TextField "Label_A_Bits" at 454,196 size 108x16; Text 'A_Bits'
   Slider "V_Range" at 566,4 size 60x160; Caption 'SIMATIC'
      Visibility <- "D_Range"
   TextField "Label_V_Range" at 566,196 size 108x16; Text 'V_Range'
   Slider "V_Bit" at 678,4 size 60x160; Caption 'SIMATIC'
      Visibility <- "D_Vis"
   TextField "Label_V_Bit" at 678,196 size 108x16; Text 'V_Bit'
   Slider "M_H" at 6,216 size 60x160; Caption 'SIMATIC'
      HorizontalMovement <- "D_Pct"
   TextField "Label_M_H" at 6,408 size 108x16; Text 'M_H'
   Slider "M_V" at 118,216 size 60x160; Caption 'SIMATIC'
      VerticalMovement <- "D_Pct"
   TextField "Label_M_V" at 118,408 size 108x16; Text 'M_V'
   Slider "M_D" at 230,216 size 60x160; Caption 'SIMATIC'
      DiagonalMovement <- "D_Pct"
   TextField "Label_M_D" at 230,408 size 108x16; Text 'M_D'
   Slider "M_Direct" at 342,216 size 60x160; Caption 'SIMATIC'
      DirectMovement <- "D_X"
      DirectMovement <- "D_Y"
   TextField "Label_M_Direct" at 342,408 size 108x16; Text 'M_Direct'
   Slider "E_Range" at 454,216 size 60x160; Caption 'SIMATIC'
      ObjectEnable <- "D_Range"
   TextField "Label_E_Range" at 454,408 size 108x16; Text 'E_Range'
   Slider "E_Bit" at 566,216 size 60x160; Caption 'SIMATIC'
      ObjectEnable <- "D_En"
   TextField "Label_E_Bit" at 566,408 size 108x16; Text 'E_Bit'
   Slider "PV_Pct" at 678,216 size 60x160; Caption 'SIMATIC'
      ProcessValue <- "D_Pct"
   TextField "Label_PV_Pct" at 678,408 size 108x16; Text 'PV_Pct'
   IOField "State" at 4,454 size 60x22; FormatPattern 9
      ProcessValue <- "D_State"
   Button "S1" at 70,454 size 40x22; TextOff 'S1'
      on Click: "SetS1"()
   Button "S2" at 114,454 size 40x22; TextOff 'S2'
      on Click: "SetS2"()
   Button "S3" at 158,454 size 40x22; TextOff 'S3'
      on Click: "SetS3"()
   Button "S4" at 202,454 size 40x22; TextOff 'S4'
      on Click: "SetS4"()
   Button "Next" at 756,454 size 40x22; TextOff 'Next'
      on Click: ActivateScreen("D_Slider_2", 0)

screen "D_Slider_2" 800x480
   Slider "PV_Int" at 6,4 size 60x160; Caption 'SIMATIC'
      ProcessValue <- "D_Int"
   TextField "Label_PV_Int" at 6,196 size 108x16; Text 'PV_Int'
   Slider "PV_Pct_0_200" at 118,4 size 60x160; Caption 'SIMATIC'
      ProcessValue <- "D_Pct"
   TextField "Label_PV_Pct_0_200" at 118,196 size 108x16; Text 'PV_Pct_0_200'
   IOField "State" at 4,454 size 60x22; FormatPattern 9
      ProcessValue <- "D_State"
   Button "S1" at 70,454 size 40x22; TextOff 'S1'
      on Click: "SetS1"()
   Button "S2" at 114,454 size 40x22; TextOff 'S2'
      on Click: "SetS2"()
   Button "S3" at 158,454 size 40x22; TextOff 'S3'
      on Click: "SetS3"()
   Button "S4" at 202,454 size 40x22; TextOff 'S4'
      on Click: "SetS4"()
   Button "Next" at 756,454 size 40x22; TextOff 'Next'
      on Click: ActivateScreen("D_Gauge_1", 0)

screen "D_SymbolLibrary_1" 800x480
   SymbolLibrary "Static" at 6,4 size 60x60
   TextField "Label_Static" at 6,96 size 108x16; Text 'Static'
   SymbolLibrary "A_Range" at 118,4 size 60x60
      Appearance <- "D_Range"
   TextField "Label_A_Range" at 118,96 size 108x16; Text 'A_Range'
   SymbolLibrary "A_Flash" at 230,4 size 60x60
      Appearance <- "D_Range"
   TextField "Label_A_Flash" at 230,96 size 108x16; Text 'A_Flash'
   SymbolLibrary "A_Bit" at 342,4 size 60x60
      Appearance <- "D_Bool"
   TextField "Label_A_Bit" at 342,96 size 108x16; Text 'A_Bit'
   SymbolLibrary "A_Bits" at 454,4 size 60x60
      Appearance <- "D_Bits"
   TextField "Label_A_Bits" at 454,96 size 108x16; Text 'A_Bits'
   SymbolLibrary "V_Range" at 566,4 size 60x60
      Visibility <- "D_Range"
   TextField "Label_V_Range" at 566,96 size 108x16; Text 'V_Range'
   SymbolLibrary "V_Bit" at 678,4 size 60x60
      Visibility <- "D_Vis"
   TextField "Label_V_Bit" at 678,96 size 108x16; Text 'V_Bit'
   SymbolLibrary "M_H" at 6,116 size 60x60
      HorizontalMovement <- "D_Pct"
   TextField "Label_M_H" at 6,208 size 108x16; Text 'M_H'
   SymbolLibrary "M_V" at 118,116 size 60x60
      VerticalMovement <- "D_Pct"
   TextField "Label_M_V" at 118,208 size 108x16; Text 'M_V'
   SymbolLibrary "M_D" at 230,116 size 60x60
      DiagonalMovement <- "D_Pct"
   TextField "Label_M_D" at 230,208 size 108x16; Text 'M_D'
   SymbolLibrary "M_Direct" at 342,116 size 60x60
      DirectMovement <- "D_X"
      DirectMovement <- "D_Y"
   TextField "Label_M_Direct" at 342,208 size 108x16; Text 'M_Direct'
   SymbolLibrary "E_Range" at 454,116 size 60x60
      ObjectEnable <- "D_Range"
   TextField "Label_E_Range" at 454,208 size 108x16; Text 'E_Range'
   SymbolLibrary "E_Bit" at 566,116 size 60x60
      ObjectEnable <- "D_En"
   TextField "Label_E_Bit" at 566,208 size 108x16; Text 'E_Bit'
   SymbolLibrary "PV_Pct" at 678,116 size 60x60
      ProcessValue <- "D_Pct"
   TextField "Label_PV_Pct" at 678,208 size 108x16; Text 'PV_Pct'
   IOField "State" at 4,454 size 60x22; FormatPattern 9
      ProcessValue <- "D_State"
   Button "S1" at 70,454 size 40x22; TextOff 'S1'
      on Click: "SetS1"()
   Button "S2" at 114,454 size 40x22; TextOff 'S2'
      on Click: "SetS2"()
   Button "S3" at 158,454 size 40x22; TextOff 'S3'
      on Click: "SetS3"()
   Button "S4" at 202,454 size 40x22; TextOff 'S4'
      on Click: "SetS4"()
   Button "Next" at 756,454 size 40x22; TextOff 'Next'
      on Click: ActivateScreen("D_Slider_1", 0)

VB script "SetS1"
   SmartTags("D_State") = 1
   SmartTags("D_Bool") = False
   SmartTags("D_SInt") = -128
   SmartTags("D_Int") = -32768
   SmartTags("D_DInt") = -2147483648
   SmartTags("D_USInt") = 0
   SmartTags("D_UInt") = 0
   SmartTags("D_UDInt") = 0
   SmartTags("D_Real") = -999.999
   SmartTags("D_LReal") = -0.00000015
   SmartTags("D_String") = ""
   SmartTags("D_DateTime") = DateSerial(1990, 1, 1) + TimeSerial(0, 0, 0)
   SmartTags("D_Pct") = 0
   SmartTags("D_Range") = 5
   SmartTags("D_Bits") = 1
   SmartTags("D_Vis") = False
   SmartTags("D_En") = False
   SmartTags("D_X") = 10
   SmartTags("D_Y") = 10
   SmartTags("D_Max") = 100
   SmartTags("D_Min") = 0
   SmartTags("D_TL") = -5
   SmartTags("D_BarR") = -5

VB script "SetS2"
   SmartTags("D_State") = 2
   SmartTags("D_Bool") = True
   SmartTags("D_SInt") = 12
   SmartTags("D_Int") = 1234
   SmartTags("D_DInt") = 123456
   SmartTags("D_USInt") = 200
   SmartTags("D_UInt") = 40000
   SmartTags("D_UDInt") = 3000000000
   SmartTags("D_Real") = 3.14159
   SmartTags("D_LReal") = 2.718281828
   SmartTags("D_String") = "Hello World"
   SmartTags("D_DateTime") = DateSerial(2026, 11, 22) + TimeSerial(13, 45, 30)
   SmartTags("D_Pct") = 50
   SmartTags("D_Range") = 25
   SmartTags("D_Bits") = 2
   SmartTags("D_Vis") = True
   SmartTags("D_En") = True
   SmartTags("D_X") = 200
   SmartTags("D_Y") = 120
   SmartTags("D_Max") = 200
   SmartTags("D_Min") = -100
   SmartTags("D_TL") = 5
   SmartTags("D_BarR") = 0

VB script "SetS3"
   SmartTags("D_State") = 3
   SmartTags("D_Bool") = True
   SmartTags("D_SInt") = 127
   SmartTags("D_Int") = 32767
   SmartTags("D_DInt") = 2147483647
   SmartTags("D_USInt") = 255
   SmartTags("D_UInt") = 65535
   SmartTags("D_UDInt") = 4294967295
   SmartTags("D_Real") = 123456.789
   SmartTags("D_LReal") = 1E+300
   SmartTags("D_String") = "Ünïcödé äöüß ÄÖÜ € – long text that is wider than the field 0123456789 ABCDEFGHIJ"
   SmartTags("D_DateTime") = DateSerial(2099, 12, 31) + TimeSerial(23, 59, 59)
   SmartTags("D_Pct") = 100
   SmartTags("D_Range") = 75
   SmartTags("D_Bits") = 4
   SmartTags("D_Vis") = True
   SmartTags("D_En") = False
   SmartTags("D_X") = 533
   SmartTags("D_Y") = 240
   SmartTags("D_Max") = 50
   SmartTags("D_Min") = -50
   SmartTags("D_TL") = 10
   SmartTags("D_BarR") = 5

VB script "SetS4"
   SmartTags("D_State") = 4
   SmartTags("D_Bool") = False
   SmartTags("D_SInt") = -1
   SmartTags("D_Int") = -1
   SmartTags("D_DInt") = 0
   SmartTags("D_USInt") = 1
   SmartTags("D_UInt") = 1
   SmartTags("D_UDInt") = 1
   SmartTags("D_Real") = 0.0005
   SmartTags("D_LReal") = -0.0
   SmartTags("D_String") = "äöü ÄÖÜ ß"
   SmartTags("D_DateTime") = DateSerial(1970, 1, 1) + TimeSerial(0, 0, 0)
   SmartTags("D_Pct") = 150
   SmartTags("D_Range") = 200
   SmartTags("D_Bits") = 9
   SmartTags("D_Vis") = False
   SmartTags("D_En") = True
   SmartTags("D_X") = -20
   SmartTags("D_Y") = 0
   SmartTags("D_Max") = 100
   SmartTags("D_Min") = 0
   SmartTags("D_TL") = 50
   SmartTags("D_BarR") = 2.5
*)

(* ===== HMI "HMI_RT_1" =====
system functions are stored by id; their names below are inferred from use
connection "HMI_Connection_3": ETHERNET, S7_1500_OMS

HMI tags "Default tag table"
   "Hmi_Bool" : Bool, internal
   "Hmi_Int" : Int, internal
   "Hmi_Real" : Real, internal
   "Hmi_String" : WString[254], internal
   "Ext_Bool" : Bool = PLC Plc_Bool AT %M100.0, 1 s
   "Ext_Int" : Int = PLC Plc_Int AT %MW102, 1 s
   "Ext_Real" : Real = PLC Plc_Real AT %MD104, 1 s
   "Ext_Byte" : Byte = PLC Plc_Byte AT %MB108, 1 s

HMI tags "C03_Tags"
   "D_State" : Int, internal
   "D_Bool" : Bool, internal
   "D_SInt" : SInt, internal
   "D_Int" : Int, internal
   "D_DInt" : DInt, internal
   "D_USInt" : USInt, internal
   "D_UInt" : UInt, internal
   "D_UDInt" : UDInt, internal
   "D_Real" : Real, internal
   "D_LReal" : LReal, internal
   "D_String" : WString[254], internal
   "D_DateTime" : DateTime, internal
   "D_Pct" : Int, internal
   "D_Range" : Int, internal
   "D_Bits" : Int, internal
   "D_Vis" : Bool, internal
   "D_En" : Bool, internal
   "D_X" : Int, internal
   "D_Y" : Int, internal
   "D_Max" : Real, internal
   "D_Min" : Real, internal
   "D_TL" : Int, internal
   "D_BarR" : Real, internal

text list "TL_Bit": 0 'Off (0)'; 1 'On (1)'

text list "TL_BitNo": 0 'Bit 0 set'; 1 'Bit 1 set'; 2 'Bit 2 set'; 3 'Bit 3 set'

text list "TL_Value": -100..-1 'Negative (-100..-1)'; 0 'Zero'; 1..9 'One to nine'; 10 'Ten: Ünïcödé äöüß ÄÖÜ €'; 32000 'Undefined value (default entry)'

screen "All_Objects" 1024x768
   TextField "TextField_1" at 680,10 size 100x30; Text 'Text'
   GraphicView "GraphicView_1" at 800,10 size 100x60
   IOField "IOField_1" at 10,90 size 100x30
   Button "Button_1" at 130,90 size 100x40; TextOff 'Text'
   SymbolicIOField "SymbolicIOField_1" at 250,90 size 120x30; TextOff '0'; TextOn '1'
   GraphicIOField "GraphicIOField_1" at 390,90 size 60x60
   DateTimeField "DateTimeField_1" at 470,90 size 160x30
   Bar "Bar_1" at 650,90 size 40x120
   Switch "Switch_1" at 710,90 size 120x40; CaptionText 'Switch'; TextOff '0'; TextOn '1'
   SymbolLibrary "SymbolLibrary_1" at 850,90 size 60x60
   Slider "Slider_1" at 930,90 size 60x160; Caption 'SIMATIC'
   Gauge "Gauge_1" at 10,270 size 150x150; CaptionText 'SIMATIC'
   Clock "Clock_1" at 180,270 size 150x150

screen "Ctl_01_AlarmView" 1024x768, template "Nav"
   AlarmView "Alarm view_1" at 3,3 size 600x300

screen "Ctl_02_TrendView" 1024x768, template "Nav"
   TrendView "Trend view_1" at 3,3 size 600x300

screen "Ctl_03_UserView" 1024x768, template "Nav"
   UserView "User view_1" at 3,3 size 480x240

screen "Ctl_04_HtmlBrowser" 1024x768, template "Nav"
   HTMLBrowser "HTML browser_1" at 3,3 size 192x192

screen "Ctl_05_WatchTable" 1024x768, template "Nav"
   StatusForce "Watch table_1" at 3,3 size 600x300; ToolTipText 'Text'

screen "Ctl_06_SmartClientView" 1024x768, template "Nav"
   SmartClientView "Sm@rtClient view_1" at 3,3 size 320x240

screen "Ctl_07_RecipeView" 1024x768, template "Nav"
   RecipeView "Recipe view_1" at 3,3 size 400x330

screen "Ctl_09_SysDiagView" 1024x768, template "Nav"
   SysDiagControl "System diagnostics view_1" at 3,3 size 600x300

screen "Ctl_10_MediaPlayer" 1024x768, template "Nav"
   MediaPlayer "Media Player_1" at 3,3 size 240x240

screen "Ctl_11_PlcCodeView" 1024x768, template "Nav"
   PLCCodeViewer "PLC code view_1" at 3,3 size 600x300

screen "Ctl_12_GraphOverview" 1024x768, template "Nav"
   S7GraphOverview "GRAPH overview_1" at 3,3 size 424x72

screen "Ctl_13_ProDiagOverview" 1024x768, template "Nav"
   ProDiagOverview "ProDiag overview_1" at 3,3 size 253x72

screen "Ctl_14_CriteriaAnalysisView" 1024x768, template "Nav"
   CriteriaAnalysisView "Criteria analysis view_1" at 3,3 size 460x150

screen "Ctl_15_CameraView" 1024x768, template "Nav"
   CameraControl "Camera view_1" at 3,3 size 320x240

screen "Ctl_16_PdfView" 1024x768, template "Nav"
   PDFView "PDFView_1" at 3,3 size 320x240

Template "Nav" 1024x768
   Button "Nav_01" at 994,2 size 28x22; TextOff 'Text'
      on Click: ActivateScreen("Ctl_01_AlarmView", 0)
   Button "Nav_02" at 994,28 size 28x22; TextOff 'Text'
      on Click: ActivateScreen("Ctl_02_TrendView", 0)
   Button "Nav_03" at 994,54 size 28x22; TextOff 'Text'
      on Click: ActivateScreen("Ctl_03_UserView", 0)
   Button "Nav_04" at 994,80 size 28x22; TextOff 'Text'
      on Click: ActivateScreen("Ctl_04_HtmlBrowser", 0)
   Button "Nav_05" at 994,106 size 28x22; TextOff 'Text'
      on Click: ActivateScreen("Ctl_05_WatchTable", 0)
   Button "Nav_06" at 994,132 size 28x22; TextOff 'Text'
      on Click: ActivateScreen("Ctl_06_SmartClientView", 0)
   Button "Nav_07" at 994,158 size 28x22; TextOff 'Text'
      on Click: ActivateScreen("Ctl_07_RecipeView", 0)
   Button "Nav_09" at 994,210 size 28x22; TextOff 'Text'
      on Click: ActivateScreen("Ctl_09_SysDiagView", 0)
   Button "Nav_10" at 994,236 size 28x22; TextOff 'Text'
      on Click: ActivateScreen("Ctl_10_MediaPlayer", 0)
   Button "Nav_11" at 994,262 size 28x22; TextOff 'Text'
      on Click: ActivateScreen("Ctl_11_PlcCodeView", 0)
   Button "Nav_12" at 994,288 size 28x22; TextOff 'Text'
      on Click: ActivateScreen("Ctl_12_GraphOverview", 0)
   Button "Nav_13" at 994,314 size 28x22; TextOff 'Text'
      on Click: ActivateScreen("Ctl_13_ProDiagOverview", 0)
   Button "Nav_14" at 994,340 size 28x22; TextOff 'Text'
      on Click: ActivateScreen("Ctl_14_CriteriaAnalysisView", 0)
   Button "Nav_15" at 994,366 size 28x22; TextOff 'Text'
      on Click: ActivateScreen("Ctl_15_CameraView", 0)
   Button "Nav_16" at 994,392 size 28x22; TextOff 'Text'
      on Click: ActivateScreen("Ctl_16_PdfView", 0)
   Button "Nav_17" at 994,418 size 28x22; TextOff 'Text'
      on Click: ActivateScreen("All_Objects", 0)

screen "P_Line_1" 1024x768
   TextField "Label_Default" at 10,62 size 108x16; Text 'Default'
   TextField "Label_BackColor" at 120,62 size 108x16; Text 'BackColor'
   TextField "Label_Color" at 230,62 size 108x16; Text 'Color'
   TextField "Label_EndStyle" at 340,62 size 108x16; Text 'EndStyle'
   TextField "Label_EndStyle_2" at 450,62 size 108x16; Text 'EndStyle_2'
   TextField "Label_EndStyle_3" at 560,62 size 108x16; Text 'EndStyle_3'
   TextField "Label_EndStyle_4" at 670,62 size 108x16; Text 'EndStyle_4'
   TextField "Label_EndStyle_5" at 780,62 size 108x16; Text 'EndStyle_5'
   TextField "Label_FillStyle" at 890,62 size 108x16; Text 'FillStyle'
   TextField "Label_Flashing" at 10,138 size 108x16; Text 'Flashing'
   TextField "Label_LineEndShapeStyle_2" at 120,138 size 108x16; Text 'LineEndShapeStyle_2'
   TextField "Label_LineWidth" at 230,138 size 108x16; Text 'LineWidth'
   TextField "Label_StartStyle" at 340,138 size 108x16; Text 'StartStyle'
   TextField "Label_StartStyle_2" at 450,138 size 108x16; Text 'StartStyle_2'
   TextField "Label_StartStyle_3" at 560,138 size 108x16; Text 'StartStyle_3'
   TextField "Label_StartStyle_4" at 670,138 size 108x16; Text 'StartStyle_4'
   TextField "Label_StartStyle_5" at 780,138 size 108x16; Text 'StartStyle_5'
   TextField "Label_Style" at 890,138 size 108x16; Text 'Style'
   TextField "Label_Style_2" at 10,214 size 108x16; Text 'Style_2'
   TextField "Label_Style_3" at 120,214 size 108x16; Text 'Style_3'
   TextField "Label_Style_4" at 230,214 size 108x16; Text 'Style_4'
   TextField "Label_UseDesignColorSchema" at 340,214 size 108x16; Text 'UseDesignColorSchema'
   Button "Next" at 982,744 size 40x22; TextOff 'Text'
      on Click: ActivateScreen("P_Polyline_1", 0)

screen "P_Polyline_1" 1024x768
   TextField "Label_Default" at 10,62 size 108x16; Text 'Default'
   TextField "Label_BackColor" at 120,62 size 108x16; Text 'BackColor'
   TextField "Label_Color" at 230,62 size 108x16; Text 'Color'
   TextField "Label_EndStyle" at 340,62 size 108x16; Text 'EndStyle'
   TextField "Label_EndStyle_2" at 450,62 size 108x16; Text 'EndStyle_2'
   TextField "Label_EndStyle_3" at 560,62 size 108x16; Text 'EndStyle_3'
   TextField "Label_EndStyle_4" at 670,62 size 108x16; Text 'EndStyle_4'
   TextField "Label_EndStyle_5" at 780,62 size 108x16; Text 'EndStyle_5'
   TextField "Label_FillStyle" at 890,62 size 108x16; Text 'FillStyle'
   TextField "Label_Flashing" at 10,138 size 108x16; Text 'Flashing'
   TextField "Label_LineEndShapeStyle_2" at 120,138 size 108x16; Text 'LineEndShapeStyle_2'
   TextField "Label_LineWidth" at 230,138 size 108x16; Text 'LineWidth'
   TextField "Label_StartStyle" at 340,138 size 108x16; Text 'StartStyle'
   TextField "Label_StartStyle_2" at 450,138 size 108x16; Text 'StartStyle_2'
   TextField "Label_StartStyle_3" at 560,138 size 108x16; Text 'StartStyle_3'
   TextField "Label_StartStyle_4" at 670,138 size 108x16; Text 'StartStyle_4'
   TextField "Label_StartStyle_5" at 780,138 size 108x16; Text 'StartStyle_5'
   TextField "Label_Style" at 890,138 size 108x16; Text 'Style'
   TextField "Label_Style_2" at 10,214 size 108x16; Text 'Style_2'
   TextField "Label_Style_3" at 120,214 size 108x16; Text 'Style_3'
   TextField "Label_Style_4" at 230,214 size 108x16; Text 'Style_4'
   TextField "Label_UseDesignColorSchema" at 340,214 size 108x16; Text 'UseDesignColorSchema'
   Button "Next" at 982,744 size 40x22; TextOff 'Text'
      on Click: ActivateScreen("P_Polygon_1", 0)

screen "P_Polygon_1" 1024x768
   TextField "Label_Default" at 10,62 size 108x16; Text 'Default'
   TextField "Label_BackColor" at 120,62 size 108x16; Text 'BackColor'
   TextField "Label_BackFillStyle" at 230,62 size 108x16; Text 'BackFillStyle'
   TextField "Label_BorderColor" at 340,62 size 108x16; Text 'BorderColor'
   TextField "Label_BorderWidth" at 450,62 size 108x16; Text 'BorderWidth'
   TextField "Label_EdgeStyle" at 560,62 size 108x16; Text 'EdgeStyle'
   TextField "Label_EdgeStyle_2" at 670,62 size 108x16; Text 'EdgeStyle_2'
   TextField "Label_EdgeStyle_3" at 780,62 size 108x16; Text 'EdgeStyle_3'
   TextField "Label_EdgeStyle_4" at 890,62 size 108x16; Text 'EdgeStyle_4'
   TextField "Label_Flashing" at 10,138 size 108x16; Text 'Flashing'
   TextField "Label_UseDesignColorSchema" at 120,138 size 108x16; Text 'UseDesignColorSchema'
   Button "Next" at 982,744 size 40x22; TextOff 'Text'
      on Click: ActivateScreen("P_Ellipse_1", 0)

screen "P_Ellipse_1" 1024x768
   TextField "Label_Default" at 10,62 size 108x16; Text 'Default'
   TextField "Label_BackColor" at 120,62 size 108x16; Text 'BackColor'
   TextField "Label_BackFillStyle" at 230,62 size 108x16; Text 'BackFillStyle'
   TextField "Label_BorderColor" at 340,62 size 108x16; Text 'BorderColor'
   TextField "Label_BorderWidth" at 450,62 size 108x16; Text 'BorderWidth'
   TextField "Label_EdgeStyle" at 560,62 size 108x16; Text 'EdgeStyle'
   TextField "Label_EdgeStyle_2" at 670,62 size 108x16; Text 'EdgeStyle_2'
   TextField "Label_EdgeStyle_3" at 780,62 size 108x16; Text 'EdgeStyle_3'
   TextField "Label_EdgeStyle_4" at 890,62 size 108x16; Text 'EdgeStyle_4'
   TextField "Label_Flashing" at 10,138 size 108x16; Text 'Flashing'
   TextField "Label_UseDesignColorSchema" at 120,138 size 108x16; Text 'UseDesignColorSchema'
   Button "Next" at 982,744 size 40x22; TextOff 'Text'
      on Click: ActivateScreen("P_Circle_1", 0)

screen "P_Circle_1" 1024x768
   TextField "Label_Default" at 10,62 size 58x16; Text 'Default'
   TextField "Label_BackColor" at 70,62 size 58x16; Text 'BackColor'
   TextField "Label_BackFillStyle" at 130,62 size 58x16; Text 'BackFillStyle'
   TextField "Label_BorderColor" at 190,62 size 58x16; Text 'BorderColor'
   TextField "Label_BorderWidth" at 250,62 size 58x16; Text 'BorderWidth'
   TextField "Label_EdgeStyle" at 310,62 size 58x16; Text 'EdgeStyle'
   TextField "Label_EdgeStyle_2" at 370,62 size 58x16; Text 'EdgeStyle_2'
   TextField "Label_EdgeStyle_3" at 430,62 size 58x16; Text 'EdgeStyle_3'
   TextField "Label_EdgeStyle_4" at 490,62 size 58x16; Text 'EdgeStyle_4'
   TextField "Label_Flashing" at 550,62 size 58x16; Text 'Flashing'
   TextField "Label_UseDesignColorSchema" at 610,62 size 58x16; Text 'UseDesignColorSchema'
   Button "Next" at 982,744 size 40x22; TextOff 'Text'
      on Click: ActivateScreen("P_Rectangle_1", 0)

screen "P_Rectangle_1" 1024x768
   TextField "Label_Default" at 10,62 size 108x16; Text 'Default'
   TextField "Label_BackColor" at 120,62 size 108x16; Text 'BackColor'
   TextField "Label_BackFillStyle" at 230,62 size 108x16; Text 'BackFillStyle'
   TextField "Label_BorderColor" at 340,62 size 108x16; Text 'BorderColor'
   TextField "Label_BorderWidth" at 450,62 size 108x16; Text 'BorderWidth'
   TextField "Label_EdgeStyle" at 560,62 size 108x16; Text 'EdgeStyle'
   TextField "Label_EdgeStyle_2" at 670,62 size 108x16; Text 'EdgeStyle_2'
   TextField "Label_EdgeStyle_3" at 780,62 size 108x16; Text 'EdgeStyle_3'
   TextField "Label_EdgeStyle_4" at 890,62 size 108x16; Text 'EdgeStyle_4'
   TextField "Label_Flashing" at 10,138 size 108x16; Text 'Flashing'
   TextField "Label_RoundCornerHeight" at 120,138 size 108x16; Text 'RoundCornerHeight'
   TextField "Label_RoundCornerWidth" at 230,138 size 108x16; Text 'RoundCornerWidth'
   TextField "Label_UseDesignColorSchema" at 340,138 size 108x16; Text 'UseDesignColorSchema'
   Button "Next" at 982,744 size 40x22; TextOff 'Text'
      on Click: ActivateScreen("P_TextField_1", 0)

screen "P_TextField_1" 1024x768
   TextField "Default" at 10,10 size 100x30; Text 'Text'
   TextField "Label_Default" at 10,42 size 108x16; Text 'Default'
   TextField "BackColor" at 120,10 size 100x30; Text 'Text'
   TextField "Label_BackColor" at 120,42 size 108x16; Text 'BackColor'
   TextField "BackFillStyle" at 230,10 size 100x30; Text 'Text'
   TextField "Label_BackFillStyle" at 230,42 size 108x16; Text 'BackFillStyle'
   TextField "BorderBackColor" at 340,10 size 100x30; Text 'Text'
   TextField "Label_BorderBackColor" at 340,42 size 108x16; Text 'BorderBackColor'
   TextField "BorderColor" at 450,10 size 100x30; Text 'Text'
   TextField "Label_BorderColor" at 450,42 size 108x16; Text 'BorderColor'
   TextField "BorderWidth" at 560,10 size 100x30; Text 'Text'
   TextField "Label_BorderWidth" at 560,42 size 108x16; Text 'BorderWidth'
   TextField "BottomMargin" at 670,10 size 100x30; Text 'Text'
   TextField "Label_BottomMargin" at 670,42 size 108x16; Text 'BottomMargin'
   TextField "CornerRadius" at 780,10 size 100x30; Text 'Text'
   TextField "Label_CornerRadius" at 780,42 size 108x16; Text 'CornerRadius'
   TextField "EdgeStyle" at 890,10 size 100x30; Text 'Text'
   TextField "Label_EdgeStyle" at 890,42 size 108x16; Text 'EdgeStyle'
   TextField "EdgeStyle_2" at 10,66 size 100x30; Text 'Text'
   TextField "Label_EdgeStyle_2" at 10,98 size 108x16; Text 'EdgeStyle_2'
   TextField "EdgeStyle_3" at 120,66 size 100x30; Text 'Text'
   TextField "Label_EdgeStyle_3" at 120,98 size 108x16; Text 'EdgeStyle_3'
   TextField "EdgeStyle_4" at 230,66 size 100x30; Text 'Text'
   TextField "Label_EdgeStyle_4" at 230,98 size 108x16; Text 'EdgeStyle_4'
   TextField "FitToLargest" at 340,66 size 100x30; Text 'Text'
   TextField "Label_FitToLargest" at 340,98 size 108x16; Text 'FitToLargest'
   TextField "Flashing" at 450,66 size 100x30; Text 'Text'
   TextField "Label_Flashing" at 450,98 size 108x16; Text 'Flashing'
   TextField "ForeColor" at 560,66 size 100x30; Text 'Text'
   TextField "Label_ForeColor" at 560,98 size 108x16; Text 'ForeColor'
   TextField "HorizontalAlignment" at 670,66 size 100x30; Text 'Text'
   TextField "Label_HorizontalAlignment" at 670,98 size 108x16; Text 'HorizontalAlignment'
   TextField "HorizontalAlignment_2" at 780,66 size 100x30; Text 'Text'
   TextField "Label_HorizontalAlignment_2" at 780,98 size 108x16; Text 'HorizontalAlignment_2'
   TextField "LeftMargin" at 890,66 size 100x30; Text 'Text'
   TextField "Label_LeftMargin" at 890,98 size 108x16; Text 'LeftMargin'
   TextField "RightMargin" at 10,122 size 100x30; Text 'Text'
   TextField "Label_RightMargin" at 10,154 size 108x16; Text 'RightMargin'
   TextField "TopMargin" at 120,122 size 100x30; Text 'Text'
   TextField "Label_TopMargin" at 120,154 size 108x16; Text 'TopMargin'
   TextField "UseDesignColorSchema" at 230,122 size 100x30; Text 'Text'
   TextField "Label_UseDesignColorSchema" at 230,154 size 108x16; Text 'UseDesignColorSchema'
   TextField "VerticalAlignment" at 340,122 size 100x30; Text 'Text'
   TextField "Label_VerticalAlignment" at 340,154 size 108x16; Text 'VerticalAlignment'
   TextField "VerticalAlignment_2" at 450,122 size 100x30; Text 'Text'
   TextField "Label_VerticalAlignment_2" at 450,154 size 108x16; Text 'VerticalAlignment_2'
   Button "Next" at 982,744 size 40x22; TextOff 'Text'
      on Click: ActivateScreen("P_GraphicView_1", 0)

screen "P_GraphicView_1" 1024x768
   GraphicView "Default" at 10,10 size 100x60
   TextField "Label_Default" at 10,72 size 108x16; Text 'Default'
   GraphicView "BackColor" at 120,10 size 100x60
   TextField "Label_BackColor" at 120,72 size 108x16; Text 'BackColor'
   GraphicView "BackFillStyle" at 230,10 size 100x60
   TextField "Label_BackFillStyle" at 230,72 size 108x16; Text 'BackFillStyle'
   GraphicView "BorderColor" at 340,10 size 100x60
   TextField "Label_BorderColor" at 340,72 size 108x16; Text 'BorderColor'
   GraphicView "BorderWidth" at 450,10 size 100x60
   TextField "Label_BorderWidth" at 450,72 size 108x16; Text 'BorderWidth'
   GraphicView "EdgeStyle" at 560,10 size 100x60
   TextField "Label_EdgeStyle" at 560,72 size 108x16; Text 'EdgeStyle'
   GraphicView "EdgeStyle_2" at 670,10 size 100x60
   TextField "Label_EdgeStyle_2" at 670,72 size 108x16; Text 'EdgeStyle_2'
   GraphicView "EdgeStyle_3" at 780,10 size 100x60
   TextField "Label_EdgeStyle_3" at 780,72 size 108x16; Text 'EdgeStyle_3'
   GraphicView "EdgeStyle_4" at 890,10 size 100x60
   TextField "Label_EdgeStyle_4" at 890,72 size 108x16; Text 'EdgeStyle_4'
   GraphicView "FitToLargest" at 10,96 size 100x60
   TextField "Label_FitToLargest" at 10,158 size 108x16; Text 'FitToLargest'
   GraphicView "Flashing" at 120,96 size 100x60
   TextField "Label_Flashing" at 120,158 size 108x16; Text 'Flashing'
   GraphicView "TransparentColor" at 230,96 size 100x60
   TextField "Label_TransparentColor" at 230,158 size 108x16; Text 'TransparentColor'
   GraphicView "UseTransparentColor" at 340,96 size 100x60
   TextField "Label_UseTransparentColor" at 340,158 size 108x16; Text 'UseTransparentColor'
   Button "Next" at 982,744 size 40x22; TextOff 'Text'
      on Click: ActivateScreen("P_IOField_1", 0)

screen "P_Button_1" 1024x768
   Button "Default" at 10,10 size 100x40; TextOff 'Text'
   TextField "Label_Default" at 10,52 size 108x16; Text 'Default'
   Button "BackColor" at 120,10 size 100x40; TextOff 'Text'
   TextField "Label_BackColor" at 120,52 size 108x16; Text 'BackColor'
   Button "BackFillStyle" at 230,10 size 100x40; TextOff 'Text'
   TextField "Label_BackFillStyle" at 230,52 size 108x16; Text 'BackFillStyle'
   Button "BorderBackColor" at 340,10 size 100x40; TextOff 'Text'
   TextField "Label_BorderBackColor" at 340,52 size 108x16; Text 'BorderBackColor'
   Button "BorderColor" at 450,10 size 100x40; TextOff 'Text'
   TextField "Label_BorderColor" at 450,52 size 108x16; Text 'BorderColor'
   Button "BorderWidth" at 560,10 size 100x40; TextOff 'Text'
   TextField "Label_BorderWidth" at 560,52 size 108x16; Text 'BorderWidth'
   Button "CornerRadius" at 670,10 size 100x40; TextOff 'Text'
   TextField "Label_CornerRadius" at 670,52 size 108x16; Text 'CornerRadius'
   Button "EdgeStyle" at 780,10 size 100x40; TextOff 'Text'
   TextField "Label_EdgeStyle" at 780,52 size 108x16; Text 'EdgeStyle'
   Button "EdgeStyle_2" at 890,10 size 100x40; TextOff 'Text'
   TextField "Label_EdgeStyle_2" at 890,52 size 108x16; Text 'EdgeStyle_2'
   Button "EdgeStyle_3" at 10,76 size 100x40; TextOff 'Text'
   TextField "Label_EdgeStyle_3" at 10,118 size 108x16; Text 'EdgeStyle_3'
   Button "EdgeStyle_4" at 120,76 size 100x40; TextOff 'Text'
   TextField "Label_EdgeStyle_4" at 120,118 size 108x16; Text 'EdgeStyle_4'
   Button "FirstGradientColor" at 230,76 size 100x40; TextOff 'Text'
   TextField "Label_FirstGradientColor" at 230,118 size 108x16; Text 'FirstGradientColor'
   Button "FirstGradientOffset" at 340,76 size 100x40; TextOff 'Text'
   TextField "Label_FirstGradientOffset" at 340,118 size 108x16; Text 'FirstGradientOffset'
   Button "FitToLargest" at 450,76 size 100x40; TextOff 'Text'
   TextField "Label_FitToLargest" at 450,118 size 108x16; Text 'FitToLargest'
   Button "Flashing" at 560,76 size 100x40; TextOff 'Text'
   TextField "Label_Flashing" at 560,118 size 108x16; Text 'Flashing'
   Button "FocusColor" at 670,76 size 100x40; TextOff 'Text'
   TextField "Label_FocusColor" at 670,118 size 108x16; Text 'FocusColor'
   Button "FocusWidth" at 780,76 size 100x40; TextOff 'Text'
   TextField "Label_FocusWidth" at 780,118 size 108x16; Text 'FocusWidth'
   Button "ForeColor" at 890,76 size 100x40; TextOff 'Text'
   TextField "Label_ForeColor" at 890,118 size 108x16; Text 'ForeColor'
   Button "HorizontalAlignment" at 10,142 size 100x40; TextOff 'Text'
   TextField "Label_HorizontalAlignment" at 10,184 size 108x16; Text 'HorizontalAlignment'
   Button "HorizontalAlignment_2" at 120,142 size 100x40; TextOff 'Text'
   TextField "Label_HorizontalAlignment_2" at 120,184 size 108x16; Text 'HorizontalAlignment_2'
   Button "HorizontalPictureAlignment" at 230,142 size 100x40; TextOff 'Text'
   TextField "Label_HorizontalPictureAlignment" at 230,184 size 108x16; Text 'HorizontalPictureAlignment'
   Button "HorizontalPictureAlignment_2" at 340,142 size 100x40; TextOff 'Text'
   TextField "Label_HorizontalPictureAlignment_2" at 340,184 size 108x16; Text 'HorizontalPictureAlignment_2'
   Button "MiddleGradientColor" at 450,142 size 100x40; TextOff 'Text'
   TextField "Label_MiddleGradientColor" at 450,184 size 108x16; Text 'MiddleGradientColor'
   Button "Mode_5" at 560,142 size 100x40; TextOff 'Text'
   TextField "Label_Mode_5" at 560,184 size 108x16; Text 'Mode_5'
   Button "Mode_7" at 670,142 size 100x40; TextOff 'Text'
   TextField "Label_Mode_7" at 670,184 size 108x16; Text 'Mode_7'
   Button "PictureAreaBottomMargin" at 780,142 size 100x40; TextOff 'Text'
   TextField "Label_PictureAreaBottomMargin" at 780,184 size 108x16; Text 'PictureAreaBottomMargin'
   Button "PictureAreaLeftMargin" at 890,142 size 100x40; TextOff 'Text'
   TextField "Label_PictureAreaLeftMargin" at 890,184 size 108x16; Text 'PictureAreaLeftMargin'
   Button "PictureAreaRightMargin" at 10,208 size 100x40; TextOff 'Text'
   TextField "Label_PictureAreaRightMargin" at 10,250 size 108x16; Text 'PictureAreaRightMargin'
   Button "PictureAreaTopMargin" at 120,208 size 100x40; TextOff 'Text'
   TextField "Label_PictureAreaTopMargin" at 120,250 size 108x16; Text 'PictureAreaTopMargin'
   Button "SecondGradientColor" at 230,208 size 100x40; TextOff 'Text'
   TextField "Label_SecondGradientColor" at 230,250 size 108x16; Text 'SecondGradientColor'
   Button "SecondGradientOffset" at 340,208 size 100x40; TextOff 'Text'
   TextField "Label_SecondGradientOffset" at 340,250 size 108x16; Text 'SecondGradientOffset'
   Button "TextAreaBottomMargin" at 450,208 size 100x40; TextOff 'Text'
   TextField "Label_TextAreaBottomMargin" at 450,250 size 108x16; Text 'TextAreaBottomMargin'
   Button "TextAreaLeftMargin" at 560,208 size 100x40; TextOff 'Text'
   TextField "Label_TextAreaLeftMargin" at 560,250 size 108x16; Text 'TextAreaLeftMargin'
   Button "TextAreaRightMargin" at 670,208 size 100x40; TextOff 'Text'
   TextField "Label_TextAreaRightMargin" at 670,250 size 108x16; Text 'TextAreaRightMargin'
   Button "TextAreaTopMargin" at 780,208 size 100x40; TextOff 'Text'
   TextField "Label_TextAreaTopMargin" at 780,250 size 108x16; Text 'TextAreaTopMargin'
   Button "UseDesignColorSchema" at 890,208 size 100x40; TextOff 'Text'
   TextField "Label_UseDesignColorSchema" at 890,250 size 108x16; Text 'UseDesignColorSchema'
   Button "UseFirstGradient" at 10,274 size 100x40; TextOff 'Text'
   TextField "Label_UseFirstGradient" at 10,316 size 108x16; Text 'UseFirstGradient'
   Button "UseSecondGradient" at 120,274 size 100x40; TextOff 'Text'
   TextField "Label_UseSecondGradient" at 120,316 size 108x16; Text 'UseSecondGradient'
   Button "VerticalAlignment" at 230,274 size 100x40; TextOff 'Text'
   TextField "Label_VerticalAlignment" at 230,316 size 108x16; Text 'VerticalAlignment'
   Button "VerticalAlignment_2" at 340,274 size 100x40; TextOff 'Text'
   TextField "Label_VerticalAlignment_2" at 340,316 size 108x16; Text 'VerticalAlignment_2'
   Button "VerticalPictureAlignment" at 450,274 size 100x40; TextOff 'Text'
   TextField "Label_VerticalPictureAlignment" at 450,316 size 108x16; Text 'VerticalPictureAlignment'
   Button "VerticalPictureAlignment_2" at 560,274 size 100x40; TextOff 'Text'
   TextField "Label_VerticalPictureAlignment_2" at 560,316 size 108x16; Text 'VerticalPictureAlignment_2'
   Button "Next" at 982,744 size 40x22; TextOff 'Text'
      on Click: ActivateScreen("P_SymbolicIOField_1", 0)

screen "P_SymbolicIOField_1" 1024x768
   SymbolicIOField "Default" at 10,10 size 120x30; TextOff '0'; TextOn '1'
   TextField "Label_Default" at 10,42 size 128x16; Text 'Default'
   SymbolicIOField "AboveUpperLimitColor" at 140,10 size 120x30; TextOff '0'; TextOn '1'
   TextField "Label_AboveUpperLimitColor" at 140,42 size 128x16; Text 'AboveUpperLimitColor'
   SymbolicIOField "BackColor" at 270,10 size 120x30; TextOff '0'; TextOn '1'
   TextField "Label_BackColor" at 270,42 size 128x16; Text 'BackColor'
   SymbolicIOField "BackFillStyle" at 400,10 size 120x30; TextOff '0'; TextOn '1'
   TextField "Label_BackFillStyle" at 400,42 size 128x16; Text 'BackFillStyle'
   SymbolicIOField "BelowLowerLimitColor" at 530,10 size 120x30; TextOff '0'; TextOn '1'
   TextField "Label_BelowLowerLimitColor" at 530,42 size 128x16; Text 'BelowLowerLimitColor'
   SymbolicIOField "BorderBackColor" at 660,10 size 120x30; TextOff '0'; TextOn '1'
   TextField "Label_BorderBackColor" at 660,42 size 128x16; Text 'BorderBackColor'
   SymbolicIOField "BorderColor" at 790,10 size 120x30; TextOff '0'; TextOn '1'
   TextField "Label_BorderColor" at 790,42 size 128x16; Text 'BorderColor'
   SymbolicIOField "BorderWidth" at 10,66 size 120x30; TextOff '0'; TextOn '1'
   TextField "Label_BorderWidth" at 10,98 size 128x16; Text 'BorderWidth'
   SymbolicIOField "BottomMargin" at 140,66 size 120x30; TextOff '0'; TextOn '1'
   TextField "Label_BottomMargin" at 140,98 size 128x16; Text 'BottomMargin'
   SymbolicIOField "CornerRadius" at 270,66 size 120x30; TextOff '0'; TextOn '1'
   TextField "Label_CornerRadius" at 270,98 size 128x16; Text 'CornerRadius'
   SymbolicIOField "CountVisibleItems" at 400,66 size 120x30; TextOff '0'; TextOn '1'
   TextField "Label_CountVisibleItems" at 400,98 size 128x16; Text 'CountVisibleItems'
   SymbolicIOField "EdgeStyle" at 530,66 size 120x30; TextOff '0'; TextOn '1'
   TextField "Label_EdgeStyle" at 530,98 size 128x16; Text 'EdgeStyle'
   SymbolicIOField "EdgeStyle_2" at 660,66 size 120x30; TextOff '0'; TextOn '1'
   TextField "Label_EdgeStyle_2" at 660,98 size 128x16; Text 'EdgeStyle_2'
   SymbolicIOField "EdgeStyle_3" at 790,66 size 120x30; TextOff '0'; TextOn '1'
   TextField "Label_EdgeStyle_3" at 790,98 size 128x16; Text 'EdgeStyle_3'
   SymbolicIOField "EdgeStyle_4" at 10,122 size 120x30; TextOff '0'; TextOn '1'
   TextField "Label_EdgeStyle_4" at 10,154 size 128x16; Text 'EdgeStyle_4'
   SymbolicIOField "EvenRowBackColor" at 140,122 size 120x30; TextOff '0'; TextOn '1'
   TextField "Label_EvenRowBackColor" at 140,154 size 128x16; Text 'EvenRowBackColor'
   SymbolicIOField "FitToLargest" at 270,122 size 120x30; TextOff '0'; TextOn '1'
   TextField "Label_FitToLargest" at 270,154 size 128x16; Text 'FitToLargest'
   SymbolicIOField "Flashing" at 400,122 size 120x30; TextOff '0'; TextOn '1'
   TextField "Label_Flashing" at 400,154 size 128x16; Text 'Flashing'
   SymbolicIOField "FlashingOnLimitViolation" at 530,122 size 120x30; TextOff '0'; TextOn '1'
   TextField "Label_FlashingOnLimitViolation" at 530,154 size 128x16; Text 'FlashingOnLimitViolation'
   SymbolicIOField "ForeColor" at 660,122 size 120x30; TextOff '0'; TextOn '1'
   TextField "Label_ForeColor" at 660,154 size 128x16; Text 'ForeColor'
   SymbolicIOField "HorizontalAlignment" at 790,122 size 120x30; TextOff '0'; TextOn '1'
   TextField "Label_HorizontalAlignment" at 790,154 size 128x16; Text 'HorizontalAlignment'
   SymbolicIOField "HorizontalAlignment_2" at 10,178 size 120x30; TextOff '0'; TextOn '1'
   TextField "Label_HorizontalAlignment_2" at 10,210 size 128x16; Text 'HorizontalAlignment_2'
   SymbolicIOField "LeftMargin" at 140,178 size 120x30; TextOff '0'; TextOn '1'
   TextField "Label_LeftMargin" at 140,210 size 128x16; Text 'LeftMargin'
   SymbolicIOField "Mode" at 270,178 size 120x30; TextOff '0'; TextOn '1'
   TextField "Label_Mode" at 270,210 size 128x16; Text 'Mode'
   SymbolicIOField "Mode_2" at 400,178 size 120x30; TextOff '0'; TextOn '1'
   TextField "Label_Mode_2" at 400,210 size 128x16; Text 'Mode_2'
   SymbolicIOField "RightMargin" at 530,178 size 120x30; TextOff '0'; TextOn '1'
   TextField "Label_RightMargin" at 530,210 size 128x16; Text 'RightMargin'
   SymbolicIOField "SelectBackColor" at 660,178 size 120x30; TextOff '0'; TextOn '1'
   TextField "Label_SelectBackColor" at 660,210 size 128x16; Text 'SelectBackColor'
   SymbolicIOField "SelectForeColor" at 790,178 size 120x30; TextOff '0'; TextOn '1'
   TextField "Label_SelectForeColor" at 790,210 size 128x16; Text 'SelectForeColor'
   SymbolicIOField "ShowDropDownButton" at 10,234 size 120x30; TextOff '0'; TextOn '1'
   TextField "Label_ShowDropDownButton" at 10,266 size 128x16; Text 'ShowDropDownButton'
   SymbolicIOField "ShowDropDownList" at 140,234 size 120x30; TextOff '0'; TextOn '1'
   TextField "Label_ShowDropDownList" at 140,266 size 128x16; Text 'ShowDropDownList'
   SymbolicIOField "TopMargin" at 270,234 size 120x30; TextOff '0'; TextOn '1'
   TextField "Label_TopMargin" at 270,266 size 128x16; Text 'TopMargin'
   SymbolicIOField "UseDesignColorSchema" at 400,234 size 120x30; TextOff '0'; TextOn '1'
   TextField "Label_UseDesignColorSchema" at 400,266 size 128x16; Text 'UseDesignColorSchema'
   SymbolicIOField "VerticalAlignment" at 530,234 size 120x30; TextOff '0'; TextOn '1'
   TextField "Label_VerticalAlignment" at 530,266 size 128x16; Text 'VerticalAlignment'
   SymbolicIOField "VerticalAlignment_2" at 660,234 size 120x30; TextOff '0'; TextOn '1'
   TextField "Label_VerticalAlignment_2" at 660,266 size 128x16; Text 'VerticalAlignment_2'
   Button "Next" at 982,744 size 40x22; TextOff 'Text'
      on Click: ActivateScreen("P_GraphicIOField_1", 0)

screen "P_GraphicIOField_1" 1024x768
   GraphicIOField "Default" at 10,10 size 60x60
   TextField "Label_Default" at 10,72 size 68x16; Text 'Default'
   GraphicIOField "AboveUpperLimitColor" at 80,10 size 60x60
   TextField "Label_AboveUpperLimitColor" at 80,72 size 68x16; Text 'AboveUpperLimitColor'
   GraphicIOField "BackColor" at 150,10 size 60x60
   TextField "Label_BackColor" at 150,72 size 68x16; Text 'BackColor'
   GraphicIOField "BackFillStyle" at 220,10 size 60x60
   TextField "Label_BackFillStyle" at 220,72 size 68x16; Text 'BackFillStyle'
   GraphicIOField "BelowLowerLimitColor" at 290,10 size 60x60
   TextField "Label_BelowLowerLimitColor" at 290,72 size 68x16; Text 'BelowLowerLimitColor'
   GraphicIOField "BorderColor" at 360,10 size 60x60
   TextField "Label_BorderColor" at 360,72 size 68x16; Text 'BorderColor'
   GraphicIOField "BorderWidth" at 430,10 size 60x60
   TextField "Label_BorderWidth" at 430,72 size 68x16; Text 'BorderWidth'
   GraphicIOField "EdgeStyle" at 500,10 size 60x60
   TextField "Label_EdgeStyle" at 500,72 size 68x16; Text 'EdgeStyle'
   GraphicIOField "EdgeStyle_2" at 570,10 size 60x60
   TextField "Label_EdgeStyle_2" at 570,72 size 68x16; Text 'EdgeStyle_2'
   GraphicIOField "EdgeStyle_3" at 640,10 size 60x60
   TextField "Label_EdgeStyle_3" at 640,72 size 68x16; Text 'EdgeStyle_3'
   GraphicIOField "EdgeStyle_4" at 710,10 size 60x60
   TextField "Label_EdgeStyle_4" at 710,72 size 68x16; Text 'EdgeStyle_4'
   GraphicIOField "FitToLargest" at 780,10 size 60x60
   TextField "Label_FitToLargest" at 780,72 size 68x16; Text 'FitToLargest'
   GraphicIOField "Flashing" at 850,10 size 60x60
   TextField "Label_Flashing" at 850,72 size 68x16; Text 'Flashing'
   GraphicIOField "FlashingOnLimitViolation" at 920,10 size 60x60
   TextField "Label_FlashingOnLimitViolation" at 920,72 size 68x16; Text 'FlashingOnLimitViolation'
   GraphicIOField "FocusColor" at 10,96 size 60x60
   TextField "Label_FocusColor" at 10,158 size 68x16; Text 'FocusColor'
   GraphicIOField "FocusWidth" at 80,96 size 60x60
   TextField "Label_FocusWidth" at 80,158 size 68x16; Text 'FocusWidth'
   GraphicIOField "Mode" at 150,96 size 60x60
   TextField "Label_Mode" at 150,158 size 68x16; Text 'Mode'
   GraphicIOField "Mode_2" at 220,96 size 60x60
   TextField "Label_Mode_2" at 220,158 size 68x16; Text 'Mode_2'
   GraphicIOField "ScrollBarOrientation" at 290,96 size 60x60
   TextField "Label_ScrollBarOrientation" at 290,158 size 68x16; Text 'ScrollBarOrientation'
   GraphicIOField "TransparentColor" at 360,96 size 60x60
   TextField "Label_TransparentColor" at 360,158 size 68x16; Text 'TransparentColor'
   GraphicIOField "UseTransparentColor" at 430,96 size 60x60
   TextField "Label_UseTransparentColor" at 430,158 size 68x16; Text 'UseTransparentColor'
   Button "Next" at 982,744 size 40x22; TextOff 'Text'
      on Click: ActivateScreen("P_DateTimeField_1", 0)

screen "P_DateTimeField_1" 1024x768
   DateTimeField "Default" at 10,10 size 160x30
   TextField "Label_Default" at 10,42 size 168x16; Text 'Default'
   DateTimeField "BackColor" at 180,10 size 160x30
   TextField "Label_BackColor" at 180,42 size 168x16; Text 'BackColor'
   DateTimeField "BackFillStyle" at 350,10 size 160x30
   TextField "Label_BackFillStyle" at 350,42 size 168x16; Text 'BackFillStyle'
   DateTimeField "BorderBackColor" at 520,10 size 160x30
   TextField "Label_BorderBackColor" at 520,42 size 168x16; Text 'BorderBackColor'
   DateTimeField "BorderColor" at 690,10 size 160x30
   TextField "Label_BorderColor" at 690,42 size 168x16; Text 'BorderColor'
   DateTimeField "BorderWidth" at 10,66 size 160x30
   TextField "Label_BorderWidth" at 10,98 size 168x16; Text 'BorderWidth'
   DateTimeField "BottomMargin" at 180,66 size 160x30
   TextField "Label_BottomMargin" at 180,98 size 168x16; Text 'BottomMargin'
   DateTimeField "CornerRadius" at 350,66 size 160x30
   TextField "Label_CornerRadius" at 350,98 size 168x16; Text 'CornerRadius'
   DateTimeField "DisplaySystemTime" at 520,66 size 160x30
   TextField "Label_DisplaySystemTime" at 520,98 size 168x16; Text 'DisplaySystemTime'
   DateTimeField "EdgeStyle" at 690,66 size 160x30
   TextField "Label_EdgeStyle" at 690,98 size 168x16; Text 'EdgeStyle'
   DateTimeField "EdgeStyle_2" at 10,122 size 160x30
   TextField "Label_EdgeStyle_2" at 10,154 size 168x16; Text 'EdgeStyle_2'
   DateTimeField "EdgeStyle_3" at 180,122 size 160x30
   TextField "Label_EdgeStyle_3" at 180,154 size 168x16; Text 'EdgeStyle_3'
   DateTimeField "EdgeStyle_4" at 350,122 size 160x30
   TextField "Label_EdgeStyle_4" at 350,154 size 168x16; Text 'EdgeStyle_4'
   DateTimeField "FitToLargest" at 520,122 size 160x30
   TextField "Label_FitToLargest" at 520,154 size 168x16; Text 'FitToLargest'
   DateTimeField "Flashing" at 690,122 size 160x30
   TextField "Label_Flashing" at 690,154 size 168x16; Text 'Flashing'
   DateTimeField "ForeColor" at 10,178 size 160x30
   TextField "Label_ForeColor" at 10,210 size 168x16; Text 'ForeColor'
   DateTimeField "HorizontalAlignment" at 180,178 size 160x30
   TextField "Label_HorizontalAlignment" at 180,210 size 168x16; Text 'HorizontalAlignment'
   DateTimeField "HorizontalAlignment_2" at 350,178 size 160x30
   TextField "Label_HorizontalAlignment_2" at 350,210 size 168x16; Text 'HorizontalAlignment_2'
   DateTimeField "LeftMargin" at 520,178 size 160x30
   TextField "Label_LeftMargin" at 520,210 size 168x16; Text 'LeftMargin'
   DateTimeField "LongDateTimeFormat" at 690,178 size 160x30
   TextField "Label_LongDateTimeFormat" at 690,210 size 168x16; Text 'LongDateTimeFormat'
   DateTimeField "Mode_3" at 10,234 size 160x30
   TextField "Label_Mode_3" at 10,266 size 168x16; Text 'Mode_3'
   DateTimeField "RightMargin" at 180,234 size 160x30
   TextField "Label_RightMargin" at 180,266 size 168x16; Text 'RightMargin'
   DateTimeField "ShowDate" at 350,234 size 160x30
   TextField "Label_ShowDate" at 350,266 size 168x16; Text 'ShowDate'
   DateTimeField "ShowTime" at 520,234 size 160x30
   TextField "Label_ShowTime" at 520,266 size 168x16; Text 'ShowTime'
   DateTimeField "TopMargin" at 690,234 size 160x30
   TextField "Label_TopMargin" at 690,266 size 168x16; Text 'TopMargin'
   DateTimeField "UseDesignColorSchema" at 10,290 size 160x30
   TextField "Label_UseDesignColorSchema" at 10,322 size 168x16; Text 'UseDesignColorSchema'
   DateTimeField "VerticalAlignment" at 180,290 size 160x30
   TextField "Label_VerticalAlignment" at 180,322 size 168x16; Text 'VerticalAlignment'
   DateTimeField "VerticalAlignment_2" at 350,290 size 160x30
   TextField "Label_VerticalAlignment_2" at 350,322 size 168x16; Text 'VerticalAlignment_2'
   Button "Next" at 982,744 size 40x22; TextOff 'Text'
      on Click: ActivateScreen("P_Bar_1", 0)

screen "P_Bar_1" 1024x768
   Bar "Default" at 10,10 size 40x120
   TextField "Label_Default" at 10,132 size 48x16; Text 'Default'
   Bar "BackColor" at 60,10 size 40x120
   TextField "Label_BackColor" at 60,132 size 48x16; Text 'BackColor'
   Bar "BarBackColor" at 110,10 size 40x120
   TextField "Label_BarBackColor" at 110,132 size 48x16; Text 'BarBackColor'
   Bar "BarEdgeStyle" at 160,10 size 40x120
   TextField "Label_BarEdgeStyle" at 160,132 size 48x16; Text 'BarEdgeStyle'
   Bar "BarEdgeStyle_2" at 210,10 size 40x120
   TextField "Label_BarEdgeStyle_2" at 210,132 size 48x16; Text 'BarEdgeStyle_2'
   Bar "BarOrientation" at 260,10 size 40x120
   TextField "Label_BarOrientation" at 260,132 size 48x16; Text 'BarOrientation'
   Bar "BarOrientation_2" at 310,10 size 40x120
   TextField "Label_BarOrientation_2" at 310,132 size 48x16; Text 'BarOrientation_2'
   Bar "BarOrientation_3" at 360,10 size 40x120
   TextField "Label_BarOrientation_3" at 360,132 size 48x16; Text 'BarOrientation_3'
   Bar "BorderBackColor" at 410,10 size 40x120
   TextField "Label_BorderBackColor" at 410,132 size 48x16; Text 'BorderBackColor'
   Bar "BorderColor" at 460,10 size 40x120
   TextField "Label_BorderColor" at 460,132 size 48x16; Text 'BorderColor'
   Bar "BorderWidth" at 510,10 size 40x120
   TextField "Label_BorderWidth" at 510,132 size 48x16; Text 'BorderWidth'
   Bar "CornerRadius" at 560,10 size 40x120
   TextField "Label_CornerRadius" at 560,132 size 48x16; Text 'CornerRadius'
   Bar "CountSubDivisions" at 610,10 size 40x120
   TextField "Label_CountSubDivisions" at 610,132 size 48x16; Text 'CountSubDivisions'
   Bar "EdgeStyle" at 660,10 size 40x120
   TextField "Label_EdgeStyle" at 660,132 size 48x16; Text 'EdgeStyle'
   Bar "EdgeStyle_2" at 710,10 size 40x120
   TextField "Label_EdgeStyle_2" at 710,132 size 48x16; Text 'EdgeStyle_2'
   Bar "EdgeStyle_3" at 760,10 size 40x120
   TextField "Label_EdgeStyle_3" at 760,132 size 48x16; Text 'EdgeStyle_3'
   Bar "EdgeStyle_4" at 810,10 size 40x120
   TextField "Label_EdgeStyle_4" at 810,132 size 48x16; Text 'EdgeStyle_4'
   Bar "Flashing" at 860,10 size 40x120
   TextField "Label_Flashing" at 860,132 size 48x16; Text 'Flashing'
   Bar "FlashingOnLimitViolation" at 910,10 size 40x120
   TextField "Label_FlashingOnLimitViolation" at 910,132 size 48x16; Text 'FlashingOnLimitViolation'
   Bar "ForeColor" at 960,10 size 40x120
   TextField "Label_ForeColor" at 960,132 size 48x16; Text 'ForeColor'
   Bar "IntegerDigits" at 10,156 size 40x120
   TextField "Label_IntegerDigits" at 10,278 size 48x16; Text 'IntegerDigits'
   Bar "LargeTickLabelingStep" at 60,156 size 40x120
   TextField "Label_LargeTickLabelingStep" at 60,278 size 48x16; Text 'LargeTickLabelingStep'
   Bar "MaximumValue" at 110,156 size 40x120; MaximumValue 200
   TextField "Label_MaximumValue" at 110,278 size 48x16; Text 'MaximumValue'
   Bar "MinimumValue" at 160,156 size 40x120; MinimumValue -100
   TextField "Label_MinimumValue" at 160,278 size 48x16; Text 'MinimumValue'
   Bar "Precision" at 210,156 size 40x120
   TextField "Label_Precision" at 210,278 size 48x16; Text 'Precision'
   Bar "RangeLower1Color" at 260,156 size 40x120
   TextField "Label_RangeLower1Color" at 260,278 size 48x16; Text 'RangeLower1Color'
   Bar "RangeLower1Enabled" at 310,156 size 40x120
   TextField "Label_RangeLower1Enabled" at 310,278 size 48x16; Text 'RangeLower1Enabled'
   Bar "RangeLower2Color" at 360,156 size 40x120
   TextField "Label_RangeLower2Color" at 360,278 size 48x16; Text 'RangeLower2Color'
   Bar "RangeLower2Enabled" at 410,156 size 40x120
   TextField "Label_RangeLower2Enabled" at 410,278 size 48x16; Text 'RangeLower2Enabled'
   Bar "RangeNormalColor" at 460,156 size 40x120
   TextField "Label_RangeNormalColor" at 460,278 size 48x16; Text 'RangeNormalColor'
   Bar "RangeNormalEnabled" at 510,156 size 40x120
   TextField "Label_RangeNormalEnabled" at 510,278 size 48x16; Text 'RangeNormalEnabled'
   Bar "RangeUpper1Color" at 560,156 size 40x120
   TextField "Label_RangeUpper1Color" at 560,278 size 48x16; Text 'RangeUpper1Color'
   Bar "RangeUpper1Enabled" at 610,156 size 40x120
   TextField "Label_RangeUpper1Enabled" at 610,278 size 48x16; Text 'RangeUpper1Enabled'
   Bar "RangeUpper2Color" at 660,156 size 40x120
   TextField "Label_RangeUpper2Color" at 660,278 size 48x16; Text 'RangeUpper2Color'
   Bar "RangeUpper2Enabled" at 710,156 size 40x120
   TextField "Label_RangeUpper2Enabled" at 710,278 size 48x16; Text 'RangeUpper2Enabled'
   Bar "ScaleColor" at 760,156 size 40x120
   TextField "Label_ScaleColor" at 760,278 size 48x16; Text 'ScaleColor'
   Bar "ScaleGradation" at 810,156 size 40x120
   TextField "Label_ScaleGradation" at 810,278 size 48x16; Text 'ScaleGradation'
   Bar "ScaleLabelingDoubleLined" at 860,156 size 40x120
   TextField "Label_ScaleLabelingDoubleLined" at 860,278 size 48x16; Text 'ScaleLabelingDoubleLined'
   Bar "ScalePosition" at 910,156 size 40x120
   TextField "Label_ScalePosition" at 910,278 size 48x16; Text 'ScalePosition'
   Bar "SegmentColoring" at 960,156 size 40x120
   TextField "Label_SegmentColoring" at 960,278 size 48x16; Text 'SegmentColoring'
   Bar "ShowLimitLines" at 10,302 size 40x120
   TextField "Label_ShowLimitLines" at 10,424 size 48x16; Text 'ShowLimitLines'
   Bar "ShowLimitMarkers" at 60,302 size 40x120
   TextField "Label_ShowLimitMarkers" at 60,424 size 48x16; Text 'ShowLimitMarkers'
   Bar "ShowLimitRanges" at 110,302 size 40x120
   TextField "Label_ShowLimitRanges" at 110,424 size 48x16; Text 'ShowLimitRanges'
   Bar "ShowProcessValue" at 160,302 size 40x120
   TextField "Label_ShowProcessValue" at 160,424 size 48x16; Text 'ShowProcessValue'
   Bar "ShowScale" at 210,302 size 40x120
   TextField "Label_ShowScale" at 210,424 size 48x16; Text 'ShowScale'
   Bar "ShowTickLabels" at 260,302 size 40x120
   TextField "Label_ShowTickLabels" at 260,424 size 48x16; Text 'ShowTickLabels'
   Bar "Unit" at 310,302 size 40x120; Unit mm
   TextField "Label_Unit" at 310,424 size 48x16; Text 'Unit'
   Bar "UseAutoScaling" at 360,302 size 40x120
   TextField "Label_UseAutoScaling" at 360,424 size 48x16; Text 'UseAutoScaling'
   Bar "UseDesignColorSchema" at 410,302 size 40x120
   TextField "Label_UseDesignColorSchema" at 410,424 size 48x16; Text 'UseDesignColorSchema'
   Bar "UseExponentialFormat" at 460,302 size 40x120
   TextField "Label_UseExponentialFormat" at 460,424 size 48x16; Text 'UseExponentialFormat'
   Button "Next" at 982,744 size 40x22; TextOff 'Text'
      on Click: ActivateScreen("P_Switch_1", 0)

screen "P_Switch_1" 1024x768
   Switch "Default" at 10,10 size 120x40; CaptionText 'Switch'; TextOff '0'; TextOn '1'
   TextField "Label_Default" at 10,52 size 128x16; Text 'Default'
   Switch "AboveUpperLimitColor" at 140,10 size 120x40; CaptionText 'Switch'; TextOff '0'; TextOn '1'
   TextField "Label_AboveUpperLimitColor" at 140,52 size 128x16; Text 'AboveUpperLimitColor'
   Switch "BackColor" at 270,10 size 120x40; CaptionText 'Switch'; TextOff '0'; TextOn '1'
   TextField "Label_BackColor" at 270,52 size 128x16; Text 'BackColor'
   Switch "BackFillStyle" at 400,10 size 120x40; CaptionText 'Switch'; TextOff '0'; TextOn '1'
   TextField "Label_BackFillStyle" at 400,52 size 128x16; Text 'BackFillStyle'
   Switch "BelowLowerLimitColor" at 530,10 size 120x40; CaptionText 'Switch'; TextOff '0'; TextOn '1'
   TextField "Label_BelowLowerLimitColor" at 530,52 size 128x16; Text 'BelowLowerLimitColor'
   Switch "BorderBackColor" at 660,10 size 120x40; CaptionText 'Switch'; TextOff '0'; TextOn '1'
   TextField "Label_BorderBackColor" at 660,52 size 128x16; Text 'BorderBackColor'
   Switch "BorderColor" at 790,10 size 120x40; CaptionText 'Switch'; TextOff '0'; TextOn '1'
   TextField "Label_BorderColor" at 790,52 size 128x16; Text 'BorderColor'
   Switch "BorderWidth" at 10,76 size 120x40; CaptionText 'Switch'; TextOff '0'; TextOn '1'
   TextField "Label_BorderWidth" at 10,118 size 128x16; Text 'BorderWidth'
   Switch "CaptionColor" at 140,76 size 120x40; CaptionText 'Switch'; TextOff '0'; TextOn '1'
   TextField "Label_CaptionColor" at 140,118 size 128x16; Text 'CaptionColor'
   Switch "CornerRadius" at 270,76 size 120x40; CaptionText 'Switch'; TextOff '0'; TextOn '1'
   TextField "Label_CornerRadius" at 270,118 size 128x16; Text 'CornerRadius'
   Switch "EdgeStyle" at 400,76 size 120x40; CaptionText 'Switch'; TextOff '0'; TextOn '1'
   TextField "Label_EdgeStyle" at 400,118 size 128x16; Text 'EdgeStyle'
   Switch "EdgeStyle_2" at 530,76 size 120x40; CaptionText 'Switch'; TextOff '0'; TextOn '1'
   TextField "Label_EdgeStyle_2" at 530,118 size 128x16; Text 'EdgeStyle_2'
   Switch "EdgeStyle_3" at 660,76 size 120x40; CaptionText 'Switch'; TextOff '0'; TextOn '1'
   TextField "Label_EdgeStyle_3" at 660,118 size 128x16; Text 'EdgeStyle_3'
   Switch "EdgeStyle_4" at 790,76 size 120x40; CaptionText 'Switch'; TextOff '0'; TextOn '1'
   TextField "Label_EdgeStyle_4" at 790,118 size 128x16; Text 'EdgeStyle_4'
   Switch "FirstGradientColor" at 10,142 size 120x40; CaptionText 'Switch'; TextOff '0'; TextOn '1'
   TextField "Label_FirstGradientColor" at 10,184 size 128x16; Text 'FirstGradientColor'
   Switch "FirstGradientOffset" at 140,142 size 120x40; CaptionText 'Switch'; TextOff '0'; TextOn '1'
   TextField "Label_FirstGradientOffset" at 140,184 size 128x16; Text 'FirstGradientOffset'
   Switch "FitToLargest" at 270,142 size 120x40; CaptionText 'Switch'; TextOff '0'; TextOn '1'
   TextField "Label_FitToLargest" at 270,184 size 128x16; Text 'FitToLargest'
   Switch "Flashing" at 400,142 size 120x40; CaptionText 'Switch'; TextOff '0'; TextOn '1'
   TextField "Label_Flashing" at 400,184 size 128x16; Text 'Flashing'
   Switch "FlashingOnLimitViolation" at 530,142 size 120x40; CaptionText 'Switch'; TextOff '0'; TextOn '1'
   TextField "Label_FlashingOnLimitViolation" at 530,184 size 128x16; Text 'FlashingOnLimitViolation'
   Switch "FocusColor" at 660,142 size 120x40; CaptionText 'Switch'; TextOff '0'; TextOn '1'
   TextField "Label_FocusColor" at 660,184 size 128x16; Text 'FocusColor'
   Switch "FocusWidth" at 790,142 size 120x40; CaptionText 'Switch'; TextOff '0'; TextOn '1'
   TextField "Label_FocusWidth" at 790,184 size 128x16; Text 'FocusWidth'
   Switch "ForeColor" at 10,208 size 120x40; CaptionText 'Switch'; TextOff '0'; TextOn '1'
   TextField "Label_ForeColor" at 10,250 size 128x16; Text 'ForeColor'
   Switch "HorizontalAlignment" at 140,208 size 120x40; CaptionText 'Switch'; TextOff '0'; TextOn '1'
   TextField "Label_HorizontalAlignment" at 140,250 size 128x16; Text 'HorizontalAlignment'
   Switch "HorizontalAlignment_2" at 270,208 size 120x40; CaptionText 'Switch'; TextOff '0'; TextOn '1'
   TextField "Label_HorizontalAlignment_2" at 270,250 size 128x16; Text 'HorizontalAlignment_2'
   Switch "HorizontalPictureAlignment" at 400,208 size 120x40; CaptionText 'Switch'; TextOff '0'; TextOn '1'
   TextField "Label_HorizontalPictureAlignment" at 400,250 size 128x16; Text 'HorizontalPictureAlignment'
   Switch "HorizontalPictureAlignment_2" at 530,208 size 120x40; CaptionText 'Switch'; TextOff '0'; TextOn '1'
   TextField "Label_HorizontalPictureAlignment_2" at 530,250 size 128x16; Text 'HorizontalPictureAlignment_2'
   Switch "InnerBackColorOff" at 660,208 size 120x40; CaptionText 'Switch'; TextOff '0'; TextOn '1'
   TextField "Label_InnerBackColorOff" at 660,250 size 128x16; Text 'InnerBackColorOff'
   Switch "InnerBackColorOn" at 790,208 size 120x40; CaptionText 'Switch'; TextOff '0'; TextOn '1'
   TextField "Label_InnerBackColorOn" at 790,250 size 128x16; Text 'InnerBackColorOn'
   Switch "MiddleGradientColor" at 10,274 size 120x40; CaptionText 'Switch'; TextOff '0'; TextOn '1'
   TextField "Label_MiddleGradientColor" at 10,316 size 128x16; Text 'MiddleGradientColor'
   Switch "PictureAreaBottomMargin" at 140,274 size 120x40; CaptionText 'Switch'; TextOff '0'; TextOn '1'
   TextField "Label_PictureAreaBottomMargin" at 140,316 size 128x16; Text 'PictureAreaBottomMargin'
   Switch "PictureAreaLeftMargin" at 270,274 size 120x40; CaptionText 'Switch'; TextOff '0'; TextOn '1'
   TextField "Label_PictureAreaLeftMargin" at 270,316 size 128x16; Text 'PictureAreaLeftMargin'
   Switch "PictureAreaRightMargin" at 400,274 size 120x40; CaptionText 'Switch'; TextOff '0'; TextOn '1'
   TextField "Label_PictureAreaRightMargin" at 400,316 size 128x16; Text 'PictureAreaRightMargin'
   Switch "PictureAreaTopMargin" at 530,274 size 120x40; CaptionText 'Switch'; TextOff '0'; TextOn '1'
   TextField "Label_PictureAreaTopMargin" at 530,316 size 128x16; Text 'PictureAreaTopMargin'
   Switch "SecondGradientColor" at 660,274 size 120x40; CaptionText 'Switch'; TextOff '0'; TextOn '1'
   TextField "Label_SecondGradientColor" at 660,316 size 128x16; Text 'SecondGradientColor'
   Switch "SecondGradientOffset" at 790,274 size 120x40; CaptionText 'Switch'; TextOff '0'; TextOn '1'
   TextField "Label_SecondGradientOffset" at 790,316 size 128x16; Text 'SecondGradientOffset'
   Switch "ShowCaption" at 10,340 size 120x40; CaptionText 'Switch'; TextOff '0'; TextOn '1'
   TextField "Label_ShowCaption" at 10,382 size 128x16; Text 'ShowCaption'
   Switch "SwitchOrientation" at 140,340 size 120x40; CaptionText 'Switch'; TextOff '0'; TextOn '1'
   TextField "Label_SwitchOrientation" at 140,382 size 128x16; Text 'SwitchOrientation'
   Switch "SwitchOrientation_2" at 270,340 size 120x40; CaptionText 'Switch'; TextOff '0'; TextOn '1'
   TextField "Label_SwitchOrientation_2" at 270,382 size 128x16; Text 'SwitchOrientation_2'
   Switch "SwitchOrientation_3" at 400,340 size 120x40; CaptionText 'Switch'; TextOff '0'; TextOn '1'
   TextField "Label_SwitchOrientation_3" at 400,382 size 128x16; Text 'SwitchOrientation_3'
   Switch "TextAreaBottomMargin" at 530,340 size 120x40; CaptionText 'Switch'; TextOff '0'; TextOn '1'
   TextField "Label_TextAreaBottomMargin" at 530,382 size 128x16; Text 'TextAreaBottomMargin'
   Switch "TextAreaLeftMargin" at 660,340 size 120x40; CaptionText 'Switch'; TextOff '0'; TextOn '1'
   TextField "Label_TextAreaLeftMargin" at 660,382 size 128x16; Text 'TextAreaLeftMargin'
   Switch "TextAreaRightMargin" at 790,340 size 120x40; CaptionText 'Switch'; TextOff '0'; TextOn '1'
   TextField "Label_TextAreaRightMargin" at 790,382 size 128x16; Text 'TextAreaRightMargin'
   Switch "TextAreaTopMargin" at 10,406 size 120x40; CaptionText 'Switch'; TextOff '0'; TextOn '1'
   TextField "Label_TextAreaTopMargin" at 10,448 size 128x16; Text 'TextAreaTopMargin'
   Switch "UseDesignColorSchema" at 140,406 size 120x40; CaptionText 'Switch'; TextOff '0'; TextOn '1'
   TextField "Label_UseDesignColorSchema" at 140,448 size 128x16; Text 'UseDesignColorSchema'
   Switch "UseFirstGradient" at 270,406 size 120x40; CaptionText 'Switch'; TextOff '0'; TextOn '1'
   TextField "Label_UseFirstGradient" at 270,448 size 128x16; Text 'UseFirstGradient'
   Switch "UseSecondGradient" at 400,406 size 120x40; CaptionText 'Switch'; TextOff '0'; TextOn '1'
   TextField "Label_UseSecondGradient" at 400,448 size 128x16; Text 'UseSecondGradient'
   Switch "VerticalAlignment" at 530,406 size 120x40; CaptionText 'Switch'; TextOff '0'; TextOn '1'
   TextField "Label_VerticalAlignment" at 530,448 size 128x16; Text 'VerticalAlignment'
   Switch "VerticalAlignment_2" at 660,406 size 120x40; CaptionText 'Switch'; TextOff '0'; TextOn '1'
   TextField "Label_VerticalAlignment_2" at 660,448 size 128x16; Text 'VerticalAlignment_2'
   Switch "VerticalPictureAlignment" at 790,406 size 120x40; CaptionText 'Switch'; TextOff '0'; TextOn '1'
   TextField "Label_VerticalPictureAlignment" at 790,448 size 128x16; Text 'VerticalPictureAlignment'
   Switch "VerticalPictureAlignment_2" at 10,472 size 120x40; CaptionText 'Switch'; TextOff '0'; TextOn '1'
   TextField "Label_VerticalPictureAlignment_2" at 10,514 size 128x16; Text 'VerticalPictureAlignment_2'
   Button "Next" at 982,744 size 40x22; TextOff 'Text'
      on Click: ActivateScreen("P_SymbolLibrary_1", 0)

screen "P_SymbolLibrary_1" 1024x768
   SymbolLibrary "Default" at 10,10 size 60x60
   TextField "Label_Default" at 10,72 size 68x16; Text 'Default'
   SymbolLibrary "AboveUpperLimitColor" at 80,10 size 60x60
   TextField "Label_AboveUpperLimitColor" at 80,72 size 68x16; Text 'AboveUpperLimitColor'
   SymbolLibrary "BackColor" at 150,10 size 60x60
   TextField "Label_BackColor" at 150,72 size 68x16; Text 'BackColor'
   SymbolLibrary "BackFillStyle" at 220,10 size 60x60
   TextField "Label_BackFillStyle" at 220,72 size 68x16; Text 'BackFillStyle'
   SymbolLibrary "BelowLowerLimitColor" at 290,10 size 60x60
   TextField "Label_BelowLowerLimitColor" at 290,72 size 68x16; Text 'BelowLowerLimitColor'
   SymbolLibrary "BlinkColor" at 360,10 size 60x60
   TextField "Label_BlinkColor" at 360,72 size 68x16; Text 'BlinkColor'
   SymbolLibrary "FillColorMode" at 430,10 size 60x60
   TextField "Label_FillColorMode" at 430,72 size 68x16; Text 'FillColorMode'
   SymbolLibrary "FillColorMode_2" at 500,10 size 60x60
   TextField "Label_FillColorMode_2" at 500,72 size 68x16; Text 'FillColorMode_2'
   SymbolLibrary "FixedAspectRatio" at 570,10 size 60x60
   TextField "Label_FixedAspectRatio" at 570,72 size 68x16; Text 'FixedAspectRatio'
   SymbolLibrary "Flashing" at 640,10 size 60x60
   TextField "Label_Flashing" at 640,72 size 68x16; Text 'Flashing'
   SymbolLibrary "FlashingOnLimitViolation" at 710,10 size 60x60
   TextField "Label_FlashingOnLimitViolation" at 710,72 size 68x16; Text 'FlashingOnLimitViolation'
   SymbolLibrary "Flip" at 780,10 size 60x60
   TextField "Label_Flip" at 780,72 size 68x16; Text 'Flip'
   SymbolLibrary "Flip_2" at 850,10 size 60x60
   TextField "Label_Flip_2" at 850,72 size 68x16; Text 'Flip_2'
   SymbolLibrary "Flip_3" at 920,10 size 60x60
   TextField "Label_Flip_3" at 920,72 size 68x16; Text 'Flip_3'
   SymbolLibrary "ForeColor" at 10,96 size 60x60
   TextField "Label_ForeColor" at 10,158 size 68x16; Text 'ForeColor'
   SymbolLibrary "Rotation" at 80,96 size 60x60
   TextField "Label_Rotation" at 80,158 size 68x16; Text 'Rotation'
   SymbolLibrary "Rotation_2" at 150,96 size 60x60
   TextField "Label_Rotation_2" at 150,158 size 68x16; Text 'Rotation_2'
   SymbolLibrary "Rotation_3" at 220,96 size 60x60
   TextField "Label_Rotation_3" at 220,158 size 68x16; Text 'Rotation_3'
   Button "Next" at 982,744 size 40x22; TextOff 'Text'
      on Click: ActivateScreen("P_Slider_1", 0)

